REGION Network 16: Actions for STATE Num:49 Wait for Centering Slide Advance
   RUNG wire#powerrail
      Contact( #s49_WaitCentSlideAdv )
      Coil( #qCenteringSlideAdvance )
   END_RUNG
   // the same network as SCL:
   #qCenteringSlideAdvance := #s49_WaitCentSlideAdv;
END_REGION

REGION Network 17: Transition for STATE Num:50 Wait for Distance Sensor Feed Back
   RUNG wire#powerrail
      Contact( #s50_WaitDistSensorFB )
      Contact( #sSst )
      Coil( #s50_WaitDistSensorFB_T1 )
   END_RUNG
   // the same network as SCL:
   #s50_WaitDistSensorFB_T1 := #s50_WaitDistSensorFB AND #sSst;
END_REGION

REGION Network 18: STATE Num:50 Wait for Distance Sensor Feed Back
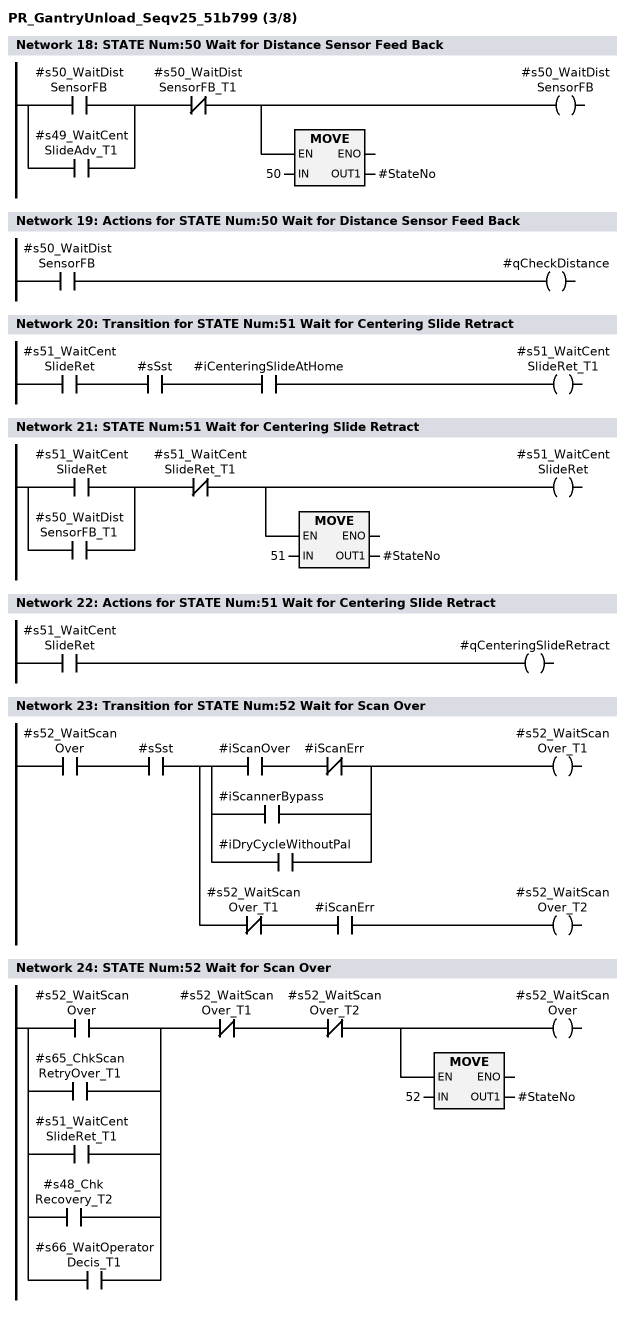
   RUNG wire#powerrail
      Contact( #s50_WaitDistSensorFB )
      wire#w1
      I_Contact( #s50_WaitDistSensorFB_T1 )
      wire#w2
      Coil( #s50_WaitDistSensorFB )
   END_RUNG
   RUNG wire#powerrail
      Contact( #s49_WaitCentSlideAdv_T1 )
   END_RUNG wire#w1
   RUNG wire#w2
      { S7_GenerateENO := "TRUE" } Move(in := 50, out1 => #StateNo)
   END_RUNG
   // the same network as SCL:
   #s50_WaitDistSensorFB := (#s50_WaitDistSensorFB OR #s49_WaitCentSlideAdv_T1) AND NOT #s50_WaitDistSensorFB_T1;
   IF #s50_WaitDistSensorFB THEN #StateNo := 50; END_IF;
END_REGION

REGION Network 19: Actions for STATE Num:50 Wait for Distance Sensor Feed Back
   RUNG wire#powerrail
      Contact( #s50_WaitDistSensorFB )
      Coil( #qCheckDistance )
   END_RUNG
   // the same network as SCL:
   #qCheckDistance := #s50_WaitDistSensorFB;
END_REGION

REGION Network 20: Transition for STATE Num:51 Wait for Centering Slide Retract
   RUNG wire#powerrail
      Contact( #s51_WaitCentSlideRet )
      Contact( #sSst )
      Contact( #iCenteringSlideAtHome )
      Coil( #s51_WaitCentSlideRet_T1 )
   END_RUNG
   // the same network as SCL:
   #s51_WaitCentSlideRet_T1 := #s51_WaitCentSlideRet AND #sSst AND #iCenteringSlideAtHome;
END_REGION

REGION Network 21: STATE Num:51 Wait for Centering Slide Retract
   RUNG wire#powerrail
      Contact( #s51_WaitCentSlideRet )
      wire#w1
      I_Contact( #s51_WaitCentSlideRet_T1 )
      wire#w2
      Coil( #s51_WaitCentSlideRet )
   END_RUNG
   RUNG wire#powerrail
      Contact( #s50_WaitDistSensorFB_T1 )
   END_RUNG wire#w1
   RUNG wire#w2
      { S7_GenerateENO := "TRUE" } Move(in := 51, out1 => #StateNo)
   END_RUNG
   // the same network as SCL:
   #s51_WaitCentSlideRet := (#s51_WaitCentSlideRet OR #s50_WaitDistSensorFB_T1) AND NOT #s51_WaitCentSlideRet_T1;
   IF #s51_WaitCentSlideRet THEN #StateNo := 51; END_IF;
END_REGION

REGION Network 22: Actions for STATE Num:51 Wait for Centering Slide Retract
   RUNG wire#powerrail
      Contact( #s51_WaitCentSlideRet )
      Coil( #qCenteringSlideRetract )
   END_RUNG
   // the same network as SCL:
   #qCenteringSlideRetract := #s51_WaitCentSlideRet;
END_REGION

REGION Network 23: Transition for STATE Num:52 Wait for Scan Over
   RUNG wire#powerrail
      Contact( #s52_WaitScanOver )
      Contact( #sSst )
      wire#w1
      Contact( #iScanOver )
      I_Contact( #iScanErr )
      wire#w2
      Coil( #s52_WaitScanOver_T1 )
   END_RUNG
   RUNG wire#w1
      Contact( #iScannerBypass )
   END_RUNG wire#w2
   RUNG wire#w1
      Contact( #iDryCycleWithoutPal )
   END_RUNG wire#w2
   RUNG wire#w1
      I_Contact( #s52_WaitScanOver_T1 )
      Contact( #iScanErr )
      Coil( #s52_WaitScanOver_T2 )
   END_RUNG
   // the same network as SCL:
   #_w1 := #s52_WaitScanOver AND #sSst;
   #s52_WaitScanOver_T1 := #_w1 AND ((#iScanOver AND NOT #iScanErr) OR #iScannerBypass OR #iDryCycleWithoutPal);
   #s52_WaitScanOver_T2 := #_w1 AND NOT #s52_WaitScanOver_T1 AND #iScanErr;
END_REGION

REGION Network 24: STATE Num:52 Wait for Scan Over
   RUNG wire#powerrail
      Contact( #s52_WaitScanOver )
      wire#w1
      I_Contact( #s52_WaitScanOver_T1 )
      I_Contact( #s52_WaitScanOver_T2 )
      wire#w2
      Coil( #s52_WaitScanOver )
   END_RUNG
   RUNG wire#powerrail
      Contact( #s65_ChkScanRetryOver_T1 )
   END_RUNG wire#w1
   RUNG wire#powerrail
      Contact( #s51_WaitCentSlideRet_T1 )
   END_RUNG wire#w1
   RUNG wire#powerrail
      Contact( #s48_ChkRecovery_T2 )
   END_RUNG wire#w1
   RUNG wire#powerrail
      Contact( #s66_WaitOperatorDecis_T1 )
   END_RUNG wire#w1
   RUNG wire#w2
      { S7_GenerateENO := "TRUE" } Move(in := 52, out1 => #StateNo)
   END_RUNG
   // the same network as SCL:
   #s52_WaitScanOver := (#s52_WaitScanOver OR #s65_ChkScanRetryOver_T1 OR #s51_WaitCentSlideRet_T1 OR #s48_ChkRecovery_T2 OR #s66_WaitOperatorDecis_T1) AND NOT #s52_WaitScanOver_T1 AND NOT #s52_WaitScanOver_T2;
   IF #s52_WaitScanOver THEN #StateNo := 52; END_IF;
END_REGION

REGION Network 25: Actions for STATE Num:52 Wait for Scan Over
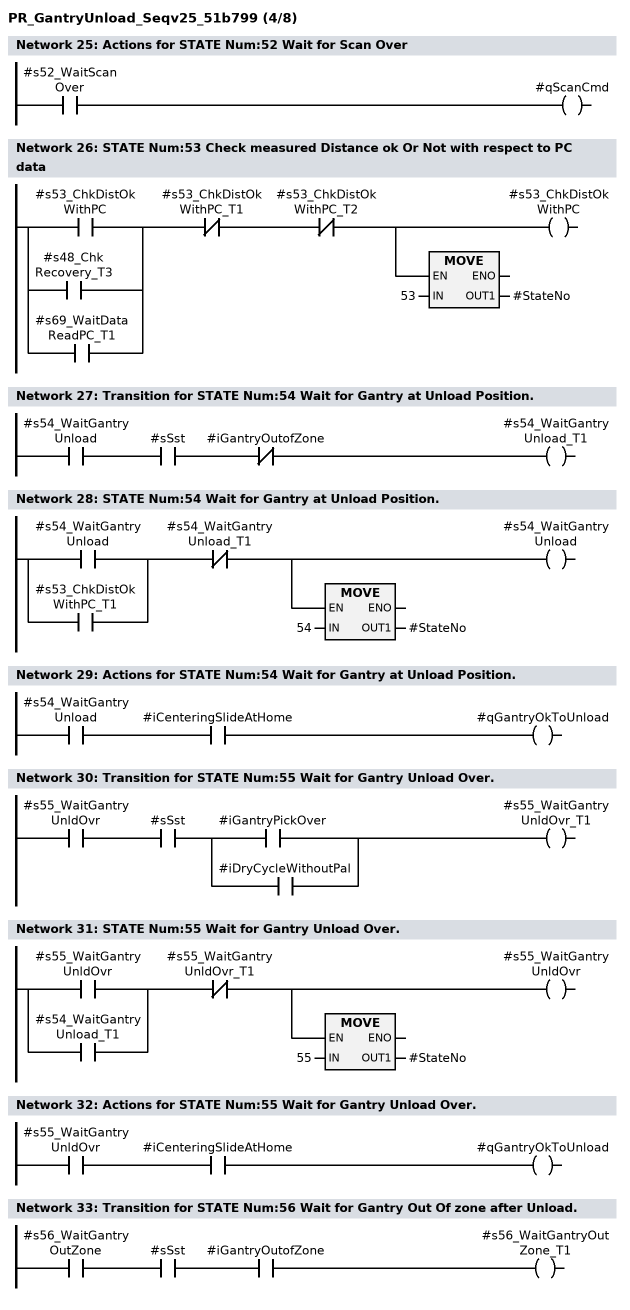
   RUNG wire#powerrail
      Contact( #s52_WaitScanOver )
      Coil( #qScanCmd )
   END_RUNG
   // the same network as SCL:
   #qScanCmd := #s52_WaitScanOver;
END_REGION

REGION Network 26: STATE Num:53 Check measured Distance ok Or Not with respect to PC data
   RUNG wire#powerrail
      Contact( #s53_ChkDistOkWithPC )
      wire#w1
      I_Contact( #s53_ChkDistOkWithPC_T1 )
      I_Contact( #s53_ChkDistOkWithPC_T2 )
      wire#w2
      Coil( #s53_ChkDistOkWithPC )
   END_RUNG
   RUNG wire#powerrail
      Contact( #s48_ChkRecovery_T3 )
   END_RUNG wire#w1
   RUNG wire#powerrail
      Contact( #s69_WaitDataReadPC_T1 )
   END_RUNG wire#w1
   RUNG wire#w2
      { S7_GenerateENO := "TRUE" } Move(in := 53, out1 => #StateNo)
   END_RUNG
   // the same network as SCL:
   #s53_ChkDistOkWithPC := (#s53_ChkDistOkWithPC OR #s48_ChkRecovery_T3 OR #s69_WaitDataReadPC_T1) AND NOT #s53_ChkDistOkWithPC_T1 AND NOT #s53_ChkDistOkWithPC_T2;
   IF #s53_ChkDistOkWithPC THEN #StateNo := 53; END_IF;
END_REGION

REGION Network 27: Transition for STATE Num:54 Wait for Gantry at Unload Position.
   RUNG wire#powerrail
      Contact( #s54_WaitGantryUnload )
      Contact( #sSst )
      I_Contact( #iGantryOutofZone )
      Coil( #s54_WaitGantryUnload_T1 )
   END_RUNG
   // the same network as SCL:
   #s54_WaitGantryUnload_T1 := #s54_WaitGantryUnload AND #sSst AND NOT #iGantryOutofZone;
END_REGION

REGION Network 28: STATE Num:54 Wait for Gantry at Unload Position.
   RUNG wire#powerrail
      Contact( #s54_WaitGantryUnload )
      wire#w1
      I_Contact( #s54_WaitGantryUnload_T1 )
      wire#w2
      Coil( #s54_WaitGantryUnload )
   END_RUNG
   RUNG wire#powerrail
      Contact( #s53_ChkDistOkWithPC_T1 )
   END_RUNG wire#w1
   RUNG wire#w2
      { S7_GenerateENO := "TRUE" } Move(in := 54, out1 => #StateNo)
   END_RUNG
   // the same network as SCL:
   #s54_WaitGantryUnload := (#s54_WaitGantryUnload OR #s53_ChkDistOkWithPC_T1) AND NOT #s54_WaitGantryUnload_T1;
   IF #s54_WaitGantryUnload THEN #StateNo := 54; END_IF;
END_REGION

REGION Network 29: Actions for STATE Num:54 Wait for Gantry at Unload Position.
   RUNG wire#powerrail
      Contact( #s54_WaitGantryUnload )
      Contact( #iCenteringSlideAtHome )
      Coil( #qGantryOkToUnload )
   END_RUNG
   // the same network as SCL:
   #qGantryOkToUnload := #s54_WaitGantryUnload AND #iCenteringSlideAtHome;
END_REGION

REGION Network 30: Transition for STATE Num:55 Wait for Gantry Unload Over.
   RUNG wire#powerrail
      Contact( #s55_WaitGantryUnldOvr )
      Contact( #sSst )
      wire#w1
      Contact( #iGantryPickOver )
      wire#w2
      Coil( #s55_WaitGantryUnldOvr_T1 )
   END_RUNG
   RUNG wire#w1
      Contact( #iDryCycleWithoutPal )
   END_RUNG wire#w2
   // the same network as SCL:
   #s55_WaitGantryUnldOvr_T1 := #s55_WaitGantryUnldOvr AND #sSst AND (#iGantryPickOver OR #iDryCycleWithoutPal);
END_REGION

REGION Network 31: STATE Num:55 Wait for Gantry Unload Over.
   RUNG wire#powerrail
      Contact( #s55_WaitGantryUnldOvr )
      wire#w1
      I_Contact( #s55_WaitGantryUnldOvr_T1 )
      wire#w2
      Coil( #s55_WaitGantryUnldOvr )
   END_RUNG
   RUNG wire#powerrail
      Contact( #s54_WaitGantryUnload_T1 )
   END_RUNG wire#w1
   RUNG wire#w2
      { S7_GenerateENO := "TRUE" } Move(in := 55, out1 => #StateNo)
   END_RUNG
   // the same network as SCL:
   #s55_WaitGantryUnldOvr := (#s55_WaitGantryUnldOvr OR #s54_WaitGantryUnload_T1) AND NOT #s55_WaitGantryUnldOvr_T1;
   IF #s55_WaitGantryUnldOvr THEN #StateNo := 55; END_IF;
END_REGION

REGION Network 32: Actions for STATE Num:55 Wait for Gantry Unload Over.
   RUNG wire#powerrail
      Contact( #s55_WaitGantryUnldOvr )
      Contact( #iCenteringSlideAtHome )
      Coil( #qGantryOkToUnload )
   END_RUNG
   // the same network as SCL:
   #qGantryOkToUnload := #s55_WaitGantryUnldOvr AND #iCenteringSlideAtHome;
END_REGION

REGION Network 33: Transition for STATE Num:56 Wait for Gantry Out Of zone after Unload.
   RUNG wire#powerrail
      Contact( #s56_WaitGantryOutZone )
      Contact( #sSst )
      Contact( #iGantryOutofZone )
      Coil( #s56_WaitGantryOutZone_T1 )
   END_RUNG
   // the same network as SCL:
   #s56_WaitGantryOutZone_T1 := #s56_WaitGantryOutZone AND #sSst AND #iGantryOutofZone;
END_REGION

REGION Network 34: STATE Num:56 Wait for Gantry Out Of zone after Unload.
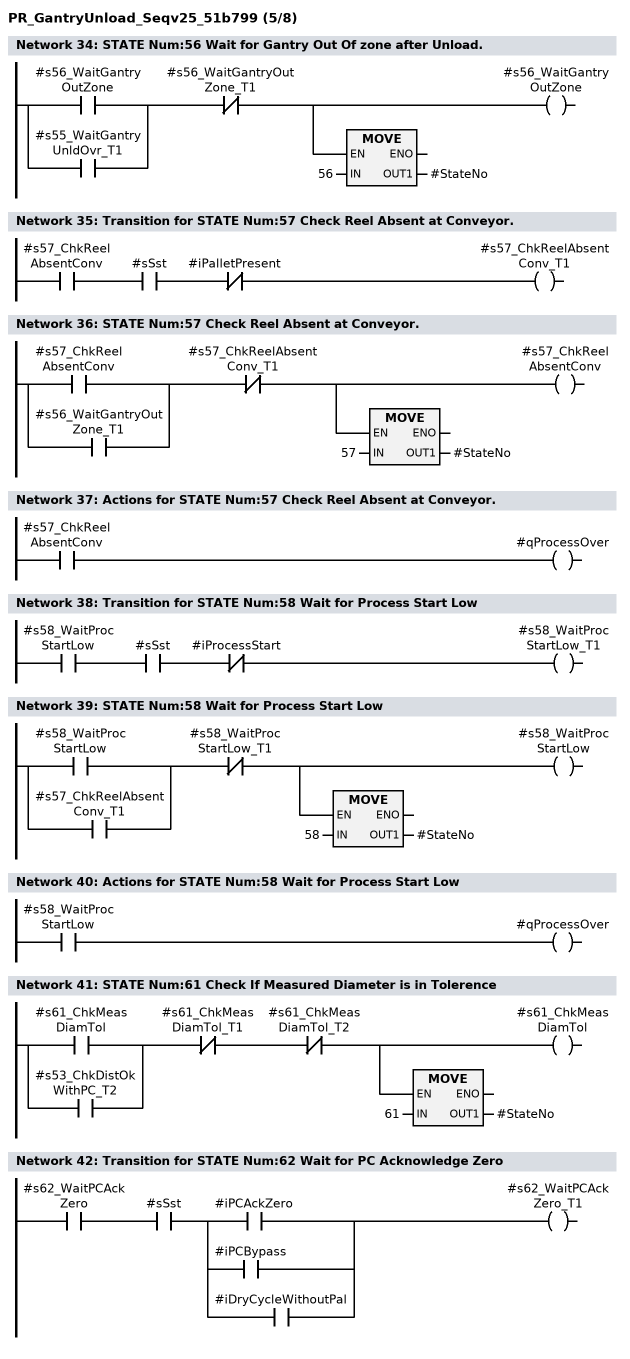
   RUNG wire#powerrail
      Contact( #s56_WaitGantryOutZone )
      wire#w1
      I_Contact( #s56_WaitGantryOutZone_T1 )
      wire#w2
      Coil( #s56_WaitGantryOutZone )
   END_RUNG
   RUNG wire#powerrail
      Contact( #s55_WaitGantryUnldOvr_T1 )
   END_RUNG wire#w1
   RUNG wire#w2
      { S7_GenerateENO := "TRUE" } Move(in := 56, out1 => #StateNo)
   END_RUNG
   // the same network as SCL:
   #s56_WaitGantryOutZone := (#s56_WaitGantryOutZone OR #s55_WaitGantryUnldOvr_T1) AND NOT #s56_WaitGantryOutZone_T1;
   IF #s56_WaitGantryOutZone THEN #StateNo := 56; END_IF;
END_REGION

REGION Network 35: Transition for STATE Num:57 Check Reel Absent at Conveyor.
   RUNG wire#powerrail
      Contact( #s57_ChkReelAbsentConv )
      Contact( #sSst )
      I_Contact( #iPalletPresent )
      Coil( #s57_ChkReelAbsentConv_T1 )
   END_RUNG
   // the same network as SCL:
   #s57_ChkReelAbsentConv_T1 := #s57_ChkReelAbsentConv AND #sSst AND NOT #iPalletPresent;
END_REGION

REGION Network 36: STATE Num:57 Check Reel Absent at Conveyor.
   RUNG wire#powerrail
      Contact( #s57_ChkReelAbsentConv )
      wire#w1
      I_Contact( #s57_ChkReelAbsentConv_T1 )
      wire#w2
      Coil( #s57_ChkReelAbsentConv )
   END_RUNG
   RUNG wire#powerrail
      Contact( #s56_WaitGantryOutZone_T1 )
   END_RUNG wire#w1
   RUNG wire#w2
      { S7_GenerateENO := "TRUE" } Move(in := 57, out1 => #StateNo)
   END_RUNG
   // the same network as SCL:
   #s57_ChkReelAbsentConv := (#s57_ChkReelAbsentConv OR #s56_WaitGantryOutZone_T1) AND NOT #s57_ChkReelAbsentConv_T1;
   IF #s57_ChkReelAbsentConv THEN #StateNo := 57; END_IF;
END_REGION

REGION Network 37: Actions for STATE Num:57 Check Reel Absent at Conveyor.
   RUNG wire#powerrail
      Contact( #s57_ChkReelAbsentConv )
      Coil( #qProcessOver )
   END_RUNG
   // the same network as SCL:
   #qProcessOver := #s57_ChkReelAbsentConv;
END_REGION

REGION Network 38: Transition for STATE Num:58 Wait for Process Start Low
   RUNG wire#powerrail
      Contact( #s58_WaitProcStartLow )
      Contact( #sSst )
      I_Contact( #iProcessStart )
      Coil( #s58_WaitProcStartLow_T1 )
   END_RUNG
   // the same network as SCL:
   #s58_WaitProcStartLow_T1 := #s58_WaitProcStartLow AND #sSst AND NOT #iProcessStart;
END_REGION

REGION Network 39: STATE Num:58 Wait for Process Start Low
   RUNG wire#powerrail
      Contact( #s58_WaitProcStartLow )
      wire#w1
      I_Contact( #s58_WaitProcStartLow_T1 )
      wire#w2
      Coil( #s58_WaitProcStartLow )
   END_RUNG
   RUNG wire#powerrail
      Contact( #s57_ChkReelAbsentConv_T1 )
   END_RUNG wire#w1
   RUNG wire#w2
      { S7_GenerateENO := "TRUE" } Move(in := 58, out1 => #StateNo)
   END_RUNG
   // the same network as SCL:
   #s58_WaitProcStartLow := (#s58_WaitProcStartLow OR #s57_ChkReelAbsentConv_T1) AND NOT #s58_WaitProcStartLow_T1;
   IF #s58_WaitProcStartLow THEN #StateNo := 58; END_IF;
END_REGION

REGION Network 40: Actions for STATE Num:58 Wait for Process Start Low
   RUNG wire#powerrail
      Contact( #s58_WaitProcStartLow )
      Coil( #qProcessOver )
   END_RUNG
   // the same network as SCL:
   #qProcessOver := #s58_WaitProcStartLow;
END_REGION

REGION Network 41: STATE Num:61 Check If Measured Diameter is in Tolerence
   RUNG wire#powerrail
      Contact( #s61_ChkMeasDiamTol )
      wire#w1
      I_Contact( #s61_ChkMeasDiamTol_T1 )
      I_Contact( #s61_ChkMeasDiamTol_T2 )
      wire#w2
      Coil( #s61_ChkMeasDiamTol )
   END_RUNG
   RUNG wire#powerrail
      Contact( #s53_ChkDistOkWithPC_T2 )
   END_RUNG wire#w1
   RUNG wire#w2
      { S7_GenerateENO := "TRUE" } Move(in := 61, out1 => #StateNo)
   END_RUNG
   // the same network as SCL:
   #s61_ChkMeasDiamTol := (#s61_ChkMeasDiamTol OR #s53_ChkDistOkWithPC_T2) AND NOT #s61_ChkMeasDiamTol_T1 AND NOT #s61_ChkMeasDiamTol_T2;
   IF #s61_ChkMeasDiamTol THEN #StateNo := 61; END_IF;
END_REGION

REGION Network 42: Transition for STATE Num:62 Wait for PC Acknowledge Zero
   RUNG wire#powerrail
      Contact( #s62_WaitPCAckZero )
      Contact( #sSst )
      wire#w1
      Contact( #iPCAckZero )
      wire#w2
      Coil( #s62_WaitPCAckZero_T1 )
   END_RUNG
   RUNG wire#w1
      Contact( #iPCBypass )
   END_RUNG wire#w2
   RUNG wire#w1
      Contact( #iDryCycleWithoutPal )
   END_RUNG wire#w2
   // the same network as SCL:
   #s62_WaitPCAckZero_T1 := #s62_WaitPCAckZero AND #sSst AND (#iPCAckZero OR #iPCBypass OR #iDryCycleWithoutPal);
END_REGION

REGION Network 43: STATE Num:62 Wait for PC Acknowledge Zero
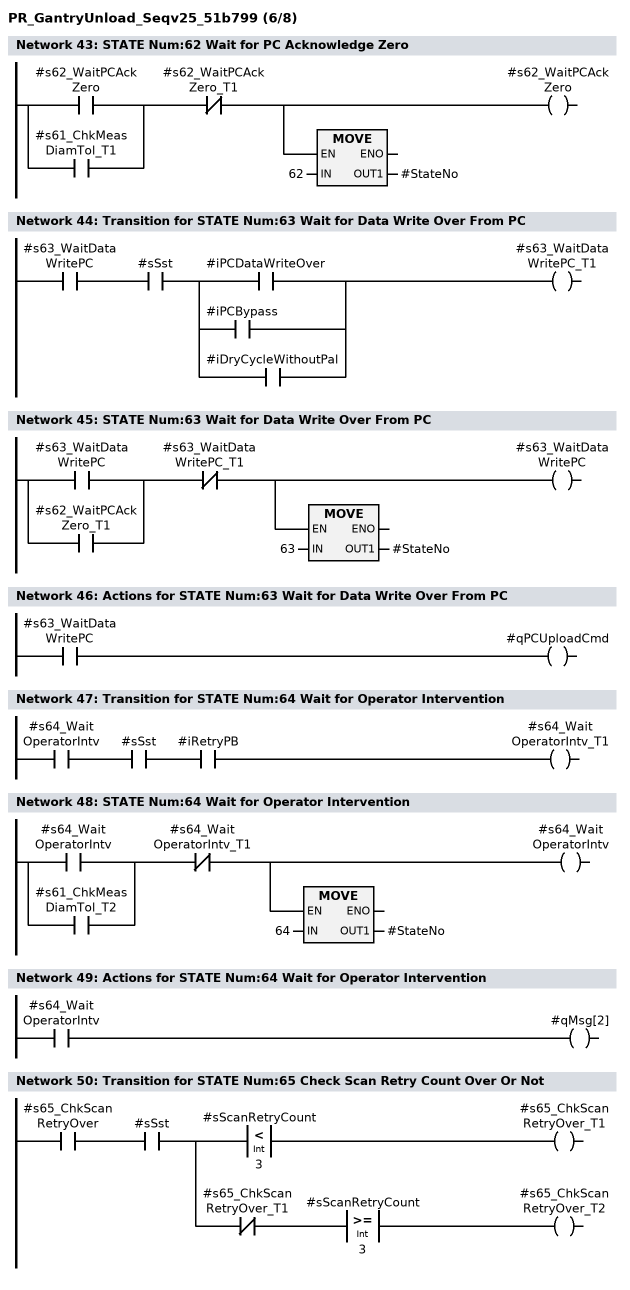
   RUNG wire#powerrail
      Contact( #s62_WaitPCAckZero )
      wire#w1
      I_Contact( #s62_WaitPCAckZero_T1 )
      wire#w2
      Coil( #s62_WaitPCAckZero )
   END_RUNG
   RUNG wire#powerrail
      Contact( #s61_ChkMeasDiamTol_T1 )
   END_RUNG wire#w1
   RUNG wire#w2
      { S7_GenerateENO := "TRUE" } Move(in := 62, out1 => #StateNo)
   END_RUNG
   // the same network as SCL:
   #s62_WaitPCAckZero := (#s62_WaitPCAckZero OR #s61_ChkMeasDiamTol_T1) AND NOT #s62_WaitPCAckZero_T1;
   IF #s62_WaitPCAckZero THEN #StateNo := 62; END_IF;
END_REGION

REGION Network 44: Transition for STATE Num:63 Wait for Data Write Over From PC
   RUNG wire#powerrail
      Contact( #s63_WaitDataWritePC )
      Contact( #sSst )
      wire#w1
      Contact( #iPCDataWriteOver )
      wire#w2
      Coil( #s63_WaitDataWritePC_T1 )
   END_RUNG
   RUNG wire#w1
      Contact( #iPCBypass )
   END_RUNG wire#w2
   RUNG wire#w1
      Contact( #iDryCycleWithoutPal )
   END_RUNG wire#w2
   // the same network as SCL:
   #s63_WaitDataWritePC_T1 := #s63_WaitDataWritePC AND #sSst AND (#iPCDataWriteOver OR #iPCBypass OR #iDryCycleWithoutPal);
END_REGION

REGION Network 45: STATE Num:63 Wait for Data Write Over From PC
   RUNG wire#powerrail
      Contact( #s63_WaitDataWritePC )
      wire#w1
      I_Contact( #s63_WaitDataWritePC_T1 )
      wire#w2
      Coil( #s63_WaitDataWritePC )
   END_RUNG
   RUNG wire#powerrail
      Contact( #s62_WaitPCAckZero_T1 )
   END_RUNG wire#w1
   RUNG wire#w2
      { S7_GenerateENO := "TRUE" } Move(in := 63, out1 => #StateNo)
   END_RUNG
   // the same network as SCL:
   #s63_WaitDataWritePC := (#s63_WaitDataWritePC OR #s62_WaitPCAckZero_T1) AND NOT #s63_WaitDataWritePC_T1;
   IF #s63_WaitDataWritePC THEN #StateNo := 63; END_IF;
END_REGION

REGION Network 46: Actions for STATE Num:63 Wait for Data Write Over From PC
   RUNG wire#powerrail
      Contact( #s63_WaitDataWritePC )
      Coil( #qPCUploadCmd )
   END_RUNG
   // the same network as SCL:
   #qPCUploadCmd := #s63_WaitDataWritePC;
END_REGION

REGION Network 47: Transition for STATE Num:64 Wait for Operator Intervention
   RUNG wire#powerrail
      Contact( #s64_WaitOperatorIntv )
      Contact( #sSst )
      Contact( #iRetryPB )
      Coil( #s64_WaitOperatorIntv_T1 )
   END_RUNG
   // the same network as SCL:
   #s64_WaitOperatorIntv_T1 := #s64_WaitOperatorIntv AND #sSst AND #iRetryPB;
END_REGION

REGION Network 48: STATE Num:64 Wait for Operator Intervention
   RUNG wire#powerrail
      Contact( #s64_WaitOperatorIntv )
      wire#w1
      I_Contact( #s64_WaitOperatorIntv_T1 )
      wire#w2
      Coil( #s64_WaitOperatorIntv )
   END_RUNG
   RUNG wire#powerrail
      Contact( #s61_ChkMeasDiamTol_T2 )
   END_RUNG wire#w1
   RUNG wire#w2
      { S7_GenerateENO := "TRUE" } Move(in := 64, out1 => #StateNo)
   END_RUNG
   // the same network as SCL:
   #s64_WaitOperatorIntv := (#s64_WaitOperatorIntv OR #s61_ChkMeasDiamTol_T2) AND NOT #s64_WaitOperatorIntv_T1;
   IF #s64_WaitOperatorIntv THEN #StateNo := 64; END_IF;
END_REGION

REGION Network 49: Actions for STATE Num:64 Wait for Operator Intervention
   RUNG wire#powerrail
      Contact( #s64_WaitOperatorIntv )
      Coil( #qMsg[2] )
   END_RUNG
   // the same network as SCL:
   #qMsg[2] := #s64_WaitOperatorIntv;
END_REGION

REGION Network 50: Transition for STATE Num:65 Check Scan Retry Count Over Or Not
   RUNG wire#powerrail
      Contact( #s65_ChkScanRetryOver )
      Contact( #sSst )
      wire#w1
      { S7_Templates := "SrcType := Int" } LT_Contact(in1 := #sScanRetryCount, in2 := 3)
      Coil( #s65_ChkScanRetryOver_T1 )
   END_RUNG
   RUNG wire#w1
      I_Contact( #s65_ChkScanRetryOver_T1 )
      { S7_Templates := "SrcType := Int" } GE_Contact(in1 := #sScanRetryCount, in2 := 3)
      Coil( #s65_ChkScanRetryOver_T2 )
   END_RUNG
   // the same network as SCL:
   #_w1 := #s65_ChkScanRetryOver AND #sSst;
   #s65_ChkScanRetryOver_T1 := #_w1 AND (#sScanRetryCount < 3);
   #s65_ChkScanRetryOver_T2 := #_w1 AND NOT #s65_ChkScanRetryOver_T1 AND (#sScanRetryCount >= 3);
END_REGION

REGION Network 51: STATE Num:65 Check Scan Retry Count Over Or Not
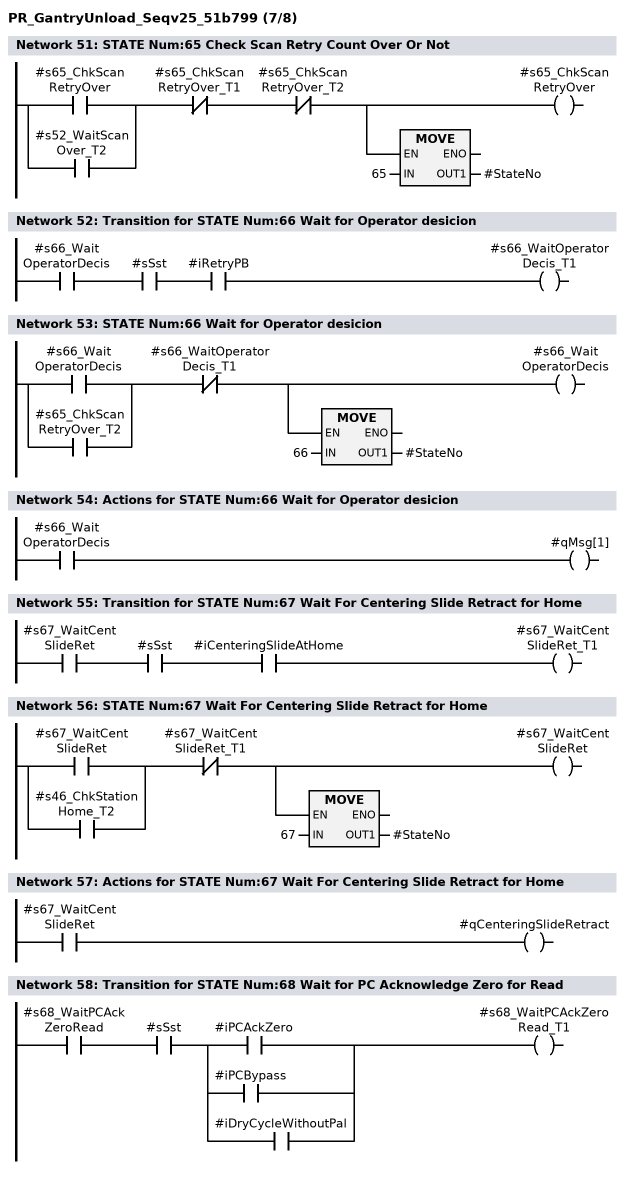
   RUNG wire#powerrail
      Contact( #s65_ChkScanRetryOver )
      wire#w1
      I_Contact( #s65_ChkScanRetryOver_T1 )
      I_Contact( #s65_ChkScanRetryOver_T2 )
      wire#w2
      Coil( #s65_ChkScanRetryOver )
   END_RUNG
   RUNG wire#powerrail
      Contact( #s52_WaitScanOver_T2 )
   END_RUNG wire#w1
   RUNG wire#w2
      { S7_GenerateENO := "TRUE" } Move(in := 65, out1 => #StateNo)
   END_RUNG
   // the same network as SCL:
   #s65_ChkScanRetryOver := (#s65_ChkScanRetryOver OR #s52_WaitScanOver_T2) AND NOT #s65_ChkScanRetryOver_T1 AND NOT #s65_ChkScanRetryOver_T2;
   IF #s65_ChkScanRetryOver THEN #StateNo := 65; END_IF;
END_REGION

REGION Network 52: Transition for STATE Num:66 Wait for Operator desicion
   RUNG wire#powerrail
      Contact( #s66_WaitOperatorDecis )
      Contact( #sSst )
      Contact( #iRetryPB )
      Coil( #s66_WaitOperatorDecis_T1 )
   END_RUNG
   // the same network as SCL:
   #s66_WaitOperatorDecis_T1 := #s66_WaitOperatorDecis AND #sSst AND #iRetryPB;
END_REGION

REGION Network 53: STATE Num:66 Wait for Operator desicion
   RUNG wire#powerrail
      Contact( #s66_WaitOperatorDecis )
      wire#w1
      I_Contact( #s66_WaitOperatorDecis_T1 )
      wire#w2
      Coil( #s66_WaitOperatorDecis )
   END_RUNG
   RUNG wire#powerrail
      Contact( #s65_ChkScanRetryOver_T2 )
   END_RUNG wire#w1
   RUNG wire#w2
      { S7_GenerateENO := "TRUE" } Move(in := 66, out1 => #StateNo)
   END_RUNG
   // the same network as SCL:
   #s66_WaitOperatorDecis := (#s66_WaitOperatorDecis OR #s65_ChkScanRetryOver_T2) AND NOT #s66_WaitOperatorDecis_T1;
   IF #s66_WaitOperatorDecis THEN #StateNo := 66; END_IF;
END_REGION

REGION Network 54: Actions for STATE Num:66 Wait for Operator desicion
   RUNG wire#powerrail
      Contact( #s66_WaitOperatorDecis )
      Coil( #qMsg[1] )
   END_RUNG
   // the same network as SCL:
   #qMsg[1] := #s66_WaitOperatorDecis;
END_REGION

REGION Network 55: Transition for STATE Num:67 Wait For Centering Slide Retract for Home
   RUNG wire#powerrail
      Contact( #s67_WaitCentSlideRet )
      Contact( #sSst )
      Contact( #iCenteringSlideAtHome )
      Coil( #s67_WaitCentSlideRet_T1 )
   END_RUNG
   // the same network as SCL:
   #s67_WaitCentSlideRet_T1 := #s67_WaitCentSlideRet AND #sSst AND #iCenteringSlideAtHome;
END_REGION

REGION Network 56: STATE Num:67 Wait For Centering Slide Retract for Home
   RUNG wire#powerrail
      Contact( #s67_WaitCentSlideRet )
      wire#w1
      I_Contact( #s67_WaitCentSlideRet_T1 )
      wire#w2
      Coil( #s67_WaitCentSlideRet )
   END_RUNG
   RUNG wire#powerrail
      Contact( #s46_ChkStationHome_T2 )
   END_RUNG wire#w1
   RUNG wire#w2
      { S7_GenerateENO := "TRUE" } Move(in := 67, out1 => #StateNo)
   END_RUNG
   // the same network as SCL:
   #s67_WaitCentSlideRet := (#s67_WaitCentSlideRet OR #s46_ChkStationHome_T2) AND NOT #s67_WaitCentSlideRet_T1;
   IF #s67_WaitCentSlideRet THEN #StateNo := 67; END_IF;
END_REGION

REGION Network 57: Actions for STATE Num:67 Wait For Centering Slide Retract for Home
   RUNG wire#powerrail
      Contact( #s67_WaitCentSlideRet )
      Coil( #qCenteringSlideRetract )
   END_RUNG
   // the same network as SCL:
   #qCenteringSlideRetract := #s67_WaitCentSlideRet;
END_REGION

REGION Network 58: Transition for STATE Num:68 Wait for PC Acknowledge Zero for Read
   RUNG wire#powerrail
      Contact( #s68_WaitPCAckZeroRead )
      Contact( #sSst )
      wire#w1
      Contact( #iPCAckZero )
      wire#w2
      Coil( #s68_WaitPCAckZeroRead_T1 )
   END_RUNG
   RUNG wire#w1
      Contact( #iPCBypass )
   END_RUNG wire#w2
   RUNG wire#w1
      Contact( #iDryCycleWithoutPal )
   END_RUNG wire#w2
   // the same network as SCL:
   #s68_WaitPCAckZeroRead_T1 := #s68_WaitPCAckZeroRead AND #sSst AND (#iPCAckZero OR #iPCBypass OR #iDryCycleWithoutPal);
END_REGION

REGION Network 59: STATE Num:68 Wait for PC Acknowledge Zero for Read
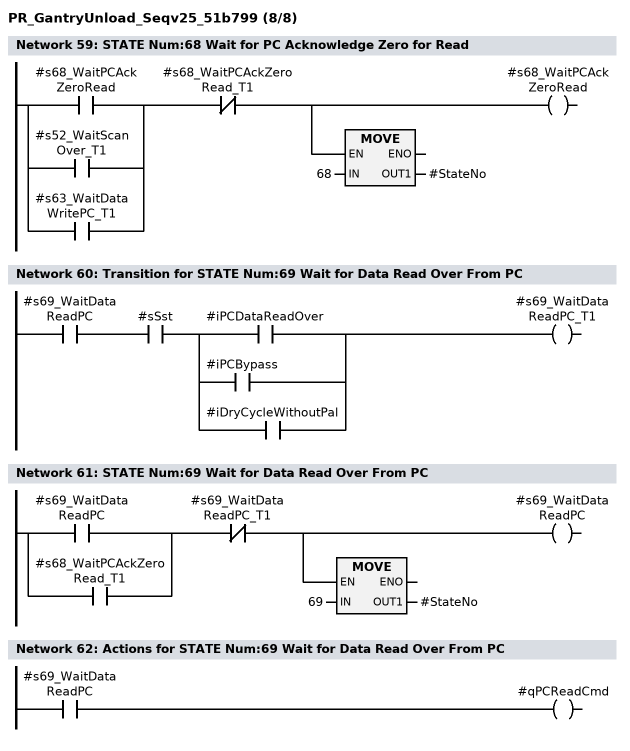
   RUNG wire#powerrail
      Contact( #s68_WaitPCAckZeroRead )
      wire#w1
      I_Contact( #s68_WaitPCAckZeroRead_T1 )
      wire#w2
      Coil( #s68_WaitPCAckZeroRead )
   END_RUNG
   RUNG wire#powerrail
      Contact( #s52_WaitScanOver_T1 )
   END_RUNG wire#w1
   RUNG wire#powerrail
      Contact( #s63_WaitDataWritePC_T1 )
   END_RUNG wire#w1
   RUNG wire#w2
      { S7_GenerateENO := "TRUE" } Move(in := 68, out1 => #StateNo)
   END_RUNG
   // the same network as SCL:
   #s68_WaitPCAckZeroRead := (#s68_WaitPCAckZeroRead OR #s52_WaitScanOver_T1 OR #s63_WaitDataWritePC_T1) AND NOT #s68_WaitPCAckZeroRead_T1;
   IF #s68_WaitPCAckZeroRead THEN #StateNo := 68; END_IF;
END_REGION

REGION Network 60: Transition for STATE Num:69 Wait for Data Read Over From PC
   RUNG wire#powerrail
      Contact( #s69_WaitDataReadPC )
      Contact( #sSst )
      wire#w1
      Contact( #iPCDataReadOver )
      wire#w2
      Coil( #s69_WaitDataReadPC_T1 )
   END_RUNG
   RUNG wire#w1
      Contact( #iPCBypass )
   END_RUNG wire#w2
   RUNG wire#w1
      Contact( #iDryCycleWithoutPal )
   END_RUNG wire#w2
   // the same network as SCL:
   #s69_WaitDataReadPC_T1 := #s69_WaitDataReadPC AND #sSst AND (#iPCDataReadOver OR #iPCBypass OR #iDryCycleWithoutPal);
END_REGION

REGION Network 61: STATE Num:69 Wait for Data Read Over From PC
   RUNG wire#powerrail
      Contact( #s69_WaitDataReadPC )
      wire#w1
      I_Contact( #s69_WaitDataReadPC_T1 )
      wire#w2
      Coil( #s69_WaitDataReadPC )
   END_RUNG
   RUNG wire#powerrail
      Contact( #s68_WaitPCAckZeroRead_T1 )
   END_RUNG wire#w1
   RUNG wire#w2
      { S7_GenerateENO := "TRUE" } Move(in := 69, out1 => #StateNo)
   END_RUNG
   // the same network as SCL:
   #s69_WaitDataReadPC := (#s69_WaitDataReadPC OR #s68_WaitPCAckZeroRead_T1) AND NOT #s69_WaitDataReadPC_T1;
   IF #s69_WaitDataReadPC THEN #StateNo := 69; END_IF;
END_REGION

REGION Network 62: Actions for STATE Num:69 Wait for Data Read Over From PC
   RUNG wire#powerrail
      Contact( #s69_WaitDataReadPC )
      Coil( #qPCReadCmd )
   END_RUNG
   // the same network as SCL:
   #qPCReadCmd := #s69_WaitDataReadPC;
END_REGION
END_FUNCTION_BLOCK

FUNCTION_BLOCK "FB_PR_GantryUnload_Seqv25_V1_V2"   // FB16, LAD
{ S7_Optimized_Access := 'TRUE' }
   VAR_INPUT
      iAutoRunning : Bool;
      iCenteringSlideAtHome : Bool;
      iCenteringSlideAtWork : Bool;
      iDistSenHighLimit : Int;
      iDistSenLowLimit : Int;
      iDistSensorIP : Int;
      iDryCycleWithoutPal : Bool;
      iGantryOutofZone : Bool;
      iGantryPickOver : Bool;
      iPCAckZero : Bool;
      iPCBypass : Bool;
      iPCDataReadOver : Bool;
      iPCDataWriteOver : Bool;
      iPalletPresent : Bool;
      iProcessStart : Bool;
      iReset_fault : Bool;
      iRetryPB : Bool;
      iScanErr : Bool;
      iScanOver : Bool;
      iScannerBypass : Bool;
      iSstMode : Bool;
      iSstPB : Bool;
   END_VAR
   VAR_OUTPUT
      qCenteringSlideAdvance : Bool;
      qCenteringSlideRetract : Bool;
      qCheckDistance : Bool;
      qGantryOkToUnload : Bool;
      qMsg : Array[0..2] of Bool;
      qPCReadCmd : Bool;
      qPCUploadCmd : Bool;
      qProcessOver : Bool;
      qScanCmd : Bool;
   END_VAR
   VAR
      StateNo : Int;
      s44_WaitResetRelease : Bool;
      s44_WaitResetRelease_T1 : Bool;
      s45_WaitGantryOutZone : Bool;
      s45_WaitGantryOutZone_T1 : Bool;
      s46_ChkStationHome : Bool;
      s46_ChkStationHome_T1 : Bool;
      s46_ChkStationHome_T2 : Bool;
      s47_WaitProcStartPZR : Bool;
      s47_WaitProcStartPZR_T1 : Bool;
      s48_ChkRecovery : Bool;
      s48_ChkRecovery_T1 : Bool;
      s48_ChkRecovery_T2 : Bool;
      s48_ChkRecovery_T3 : Bool;
      s49_WaitCentSlideAdv : Bool;
      s49_WaitCentSlideAdv_T1 : Bool;
      s50_WaitDistSensorFB : Bool;
      s50_WaitDistSensorFB_T1 : Bool;
      s51_WaitCentSlideRet : Bool;
      s51_WaitCentSlideRet_T1 : Bool;
      s52_WaitScanOver : Bool;
      s52_WaitScanOver_T1 : Bool;
      s52_WaitScanOver_T2 : Bool;
      s53_ChkMeasDistPCDat : Bool;
      s53_ChkMeasDistPCDat_T1 : Bool;
      s53_ChkMeasDistPCDat_T2 : Bool;
      s54_WaitGantryUnload : Bool;
      s54_WaitGantryUnload_T1 : Bool;
      s55_WaitGantryUnldOvr : Bool;
      s55_WaitGantryUnldOvr_T1 : Bool;
      s56_WaitGantryOutZone : Bool;
      s56_WaitGantryOutZone_T1 : Bool;
      s57_ChkReelAbsentCnv : Bool;
      s57_ChkReelAbsentCnv_T1 : Bool;
      s58_WaitProcStartLow : Bool;
      s58_WaitProcStartLow_T1 : Bool;
      s61_ChkMeasDiamTol : Bool;
      s61_ChkMeasDiamTol_T1 : Bool;
      s61_ChkMeasDiamTol_T2 : Bool;
      s62_WaitPCAckZero : Bool;
      s62_WaitPCAckZero_T1 : Bool;
      s63_WaitDataWritePC : Bool;
      s63_WaitDataWritePC_T1 : Bool;
      s64_WaitOperInterven : Bool;
      s64_WaitOperInterven_T1 : Bool;
      s65_ChkScanRetryOver : Bool;
      s65_ChkScanRetryOver_T1 : Bool;
      s65_ChkScanRetryOver_T2 : Bool;
      s66_WaitOperDecision : Bool;
      s66_WaitOperDecision_T1 : Bool;
      s67_WaitCentSlideRet : Bool;
      s67_WaitCentSlideRet_T1 : Bool;
      s68_WaitPCAckZeroRd : Bool;
      s68_WaitPCAckZeroRd_T1 : Bool;
      s69_WaitDataReadPC : Bool;
      s69_WaitDataReadPC_T1 : Bool;
      sDistanceHighLimit : Int;
      sDistanceLowLimit : Int;
      sRecoveryInt : Int;
      sScanRetryCount : Int;
      sSst : Bool;
      sSstPulse : Bool;
      sSstRise : Bool;
   END_VAR
   VAR_TEMP
      tOne : Bool;
   END_VAR
   VAR_TEMP   // added for the SCL form of the ladder/FBD networks
      _w1 : Bool;
   END_VAR
BEGIN

REGION Network 1
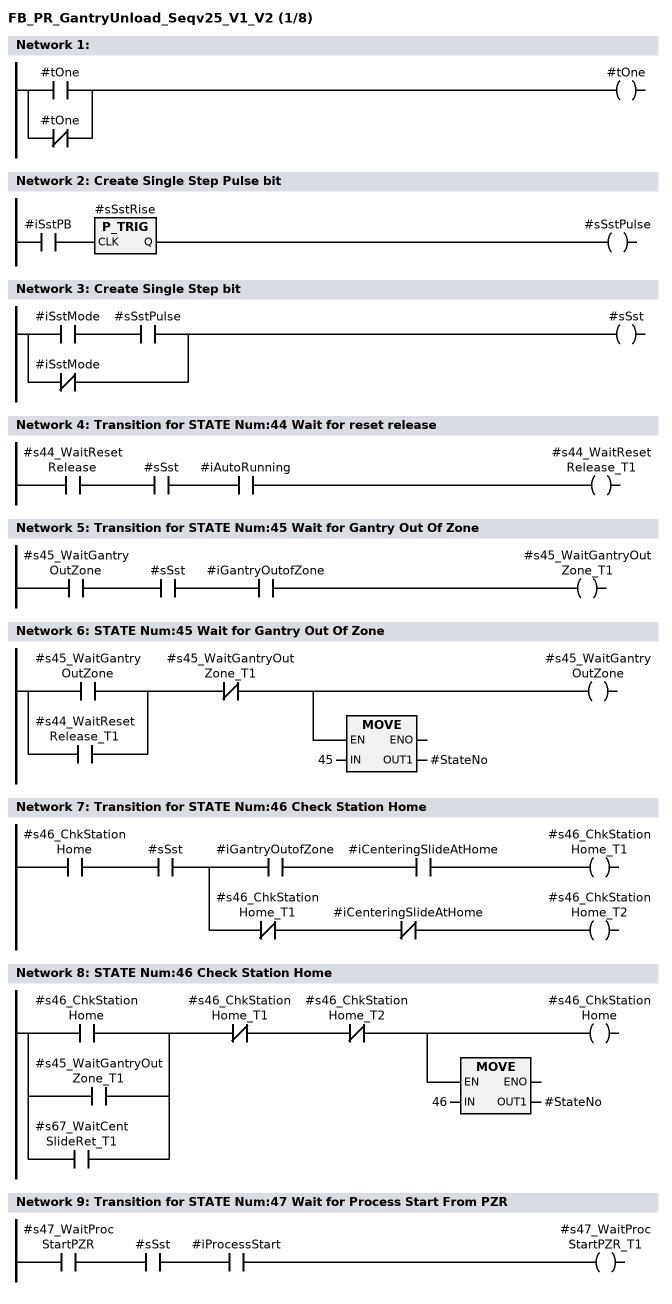
   RUNG wire#powerrail
      Contact( #tOne )
      wire#w1
      Coil( #tOne )
   END_RUNG
   RUNG wire#powerrail
      I_Contact( #tOne )
   END_RUNG wire#w1
   // the same network as SCL:
   #tOne := #tOne OR NOT #tOne;
END_REGION

REGION Network 2: Create Single Step Pulse bit
   RUNG wire#powerrail
      Contact( #iSstPB )
      P_Trig( #sSstRise )
      Coil( #sSstPulse )
   END_RUNG
   // the same network as SCL:
   #_w1 := #iSstPB AND NOT #sSstRise;   // rising edge
   #sSstRise := #iSstPB;
   #sSstPulse := #_w1;
END_REGION

REGION Network 3: Create Single Step bit
   RUNG wire#powerrail
      Contact( #iSstMode )
      Contact( #sSstPulse )
      wire#w1
      Coil( #sSst )
   END_RUNG
   RUNG wire#powerrail
      I_Contact( #iSstMode )
   END_RUNG wire#w1
   // the same network as SCL:
   #sSst := (#iSstMode AND #sSstPulse) OR NOT #iSstMode;
END_REGION

REGION Network 4: Transition for STATE Num:44 Wait for reset release
   RUNG wire#powerrail
      Contact( #s44_WaitResetRelease )
      Contact( #sSst )
      Contact( #iAutoRunning )
      Coil( #s44_WaitResetRelease_T1 )
   END_RUNG
   // the same network as SCL:
   #s44_WaitResetRelease_T1 := #s44_WaitResetRelease AND #sSst AND #iAutoRunning;
END_REGION

REGION Network 5: Transition for STATE Num:45 Wait for Gantry Out Of Zone
   RUNG wire#powerrail
      Contact( #s45_WaitGantryOutZone )
      Contact( #sSst )
      Contact( #iGantryOutofZone )
      Coil( #s45_WaitGantryOutZone_T1 )
   END_RUNG
   // the same network as SCL:
   #s45_WaitGantryOutZone_T1 := #s45_WaitGantryOutZone AND #sSst AND #iGantryOutofZone;
END_REGION

REGION Network 6: STATE Num:45 Wait for Gantry Out Of Zone
   RUNG wire#powerrail
      Contact( #s45_WaitGantryOutZone )
      wire#w1
      I_Contact( #s45_WaitGantryOutZone_T1 )
      wire#w2
      Coil( #s45_WaitGantryOutZone )
   END_RUNG
   RUNG wire#powerrail
      Contact( #s44_WaitResetRelease_T1 )
   END_RUNG wire#w1
   RUNG wire#w2
      { S7_GenerateENO := "TRUE" } Move(in := 45, out1 => #StateNo)
   END_RUNG
   // the same network as SCL:
   #s45_WaitGantryOutZone := (#s45_WaitGantryOutZone OR #s44_WaitResetRelease_T1) AND NOT #s45_WaitGantryOutZone_T1;
   IF #s45_WaitGantryOutZone THEN #StateNo := 45; END_IF;
END_REGION

REGION Network 7: Transition for STATE Num:46 Check Station Home
   RUNG wire#powerrail
      Contact( #s46_ChkStationHome )
      Contact( #sSst )
      wire#w1
      Contact( #iGantryOutofZone )
      Contact( #iCenteringSlideAtHome )
      Coil( #s46_ChkStationHome_T1 )
   END_RUNG
   RUNG wire#w1
      I_Contact( #s46_ChkStationHome_T1 )
      I_Contact( #iCenteringSlideAtHome )
      Coil( #s46_ChkStationHome_T2 )
   END_RUNG
   // the same network as SCL:
   #_w1 := #s46_ChkStationHome AND #sSst;
   #s46_ChkStationHome_T1 := #_w1 AND #iGantryOutofZone AND #iCenteringSlideAtHome;
   #s46_ChkStationHome_T2 := #_w1 AND NOT #s46_ChkStationHome_T1 AND NOT #iCenteringSlideAtHome;
END_REGION

REGION Network 8: STATE Num:46 Check Station Home
   RUNG wire#powerrail
      Contact( #s46_ChkStationHome )
      wire#w1
      I_Contact( #s46_ChkStationHome_T1 )
      I_Contact( #s46_ChkStationHome_T2 )
      wire#w2
      Coil( #s46_ChkStationHome )
   END_RUNG
   RUNG wire#powerrail
      Contact( #s45_WaitGantryOutZone_T1 )
   END_RUNG wire#w1
   RUNG wire#powerrail
      Contact( #s67_WaitCentSlideRet_T1 )
   END_RUNG wire#w1
   RUNG wire#w2
      { S7_GenerateENO := "TRUE" } Move(in := 46, out1 => #StateNo)
   END_RUNG
   // the same network as SCL:
   #s46_ChkStationHome := (#s46_ChkStationHome OR #s45_WaitGantryOutZone_T1 OR #s67_WaitCentSlideRet_T1) AND NOT #s46_ChkStationHome_T1 AND NOT #s46_ChkStationHome_T2;
   IF #s46_ChkStationHome THEN #StateNo := 46; END_IF;
END_REGION

REGION Network 9: Transition for STATE Num:47 Wait for Process Start From PZR
   RUNG wire#powerrail
      Contact( #s47_WaitProcStartPZR )
      Contact( #sSst )
      Contact( #iProcessStart )
      Coil( #s47_WaitProcStartPZR_T1 )
   END_RUNG
   // the same network as SCL:
   #s47_WaitProcStartPZR_T1 := #s47_WaitProcStartPZR AND #sSst AND #iProcessStart;
END_REGION

REGION Network 10: STATE Num:47 Wait for Process Start From PZR
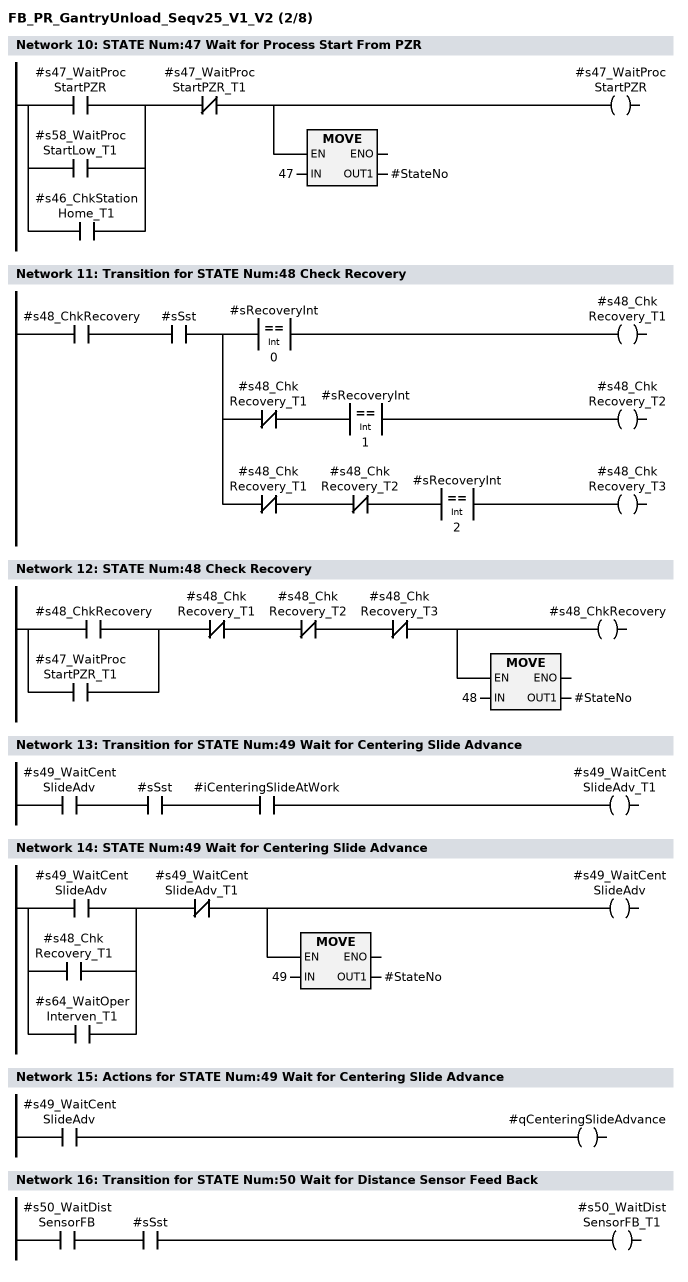
   RUNG wire#powerrail
      Contact( #s47_WaitProcStartPZR )
      wire#w1
      I_Contact( #s47_WaitProcStartPZR_T1 )
      wire#w2
      Coil( #s47_WaitProcStartPZR )
   END_RUNG
   RUNG wire#powerrail
      Contact( #s58_WaitProcStartLow_T1 )
   END_RUNG wire#w1
   RUNG wire#powerrail
      Contact( #s46_ChkStationHome_T1 )
   END_RUNG wire#w1
   RUNG wire#w2
      { S7_GenerateENO := "TRUE" } Move(in := 47, out1 => #StateNo)
   END_RUNG
   // the same network as SCL:
   #s47_WaitProcStartPZR := (#s47_WaitProcStartPZR OR #s58_WaitProcStartLow_T1 OR #s46_ChkStationHome_T1) AND NOT #s47_WaitProcStartPZR_T1;
   IF #s47_WaitProcStartPZR THEN #StateNo := 47; END_IF;
END_REGION

REGION Network 11: Transition for STATE Num:48 Check Recovery
   RUNG wire#powerrail
      Contact( #s48_ChkRecovery )
      Contact( #sSst )
      wire#w1
      { S7_Templates := "SrcType := Int" } EQ_Contact(in1 := #sRecoveryInt, in2 := 0)
      Coil( #s48_ChkRecovery_T1 )
   END_RUNG
   RUNG wire#w1
      I_Contact( #s48_ChkRecovery_T1 )
      { S7_Templates := "SrcType := Int" } EQ_Contact(in1 := #sRecoveryInt, in2 := 1)
      Coil( #s48_ChkRecovery_T2 )
   END_RUNG
   RUNG wire#w1
      I_Contact( #s48_ChkRecovery_T1 )
      I_Contact( #s48_ChkRecovery_T2 )
      { S7_Templates := "SrcType := Int" } EQ_Contact(in1 := #sRecoveryInt, in2 := 2)
      Coil( #s48_ChkRecovery_T3 )
   END_RUNG
   // the same network as SCL:
   #_w1 := #s48_ChkRecovery AND #sSst;
   #s48_ChkRecovery_T1 := #_w1 AND (#sRecoveryInt = 0);
   #s48_ChkRecovery_T2 := #_w1 AND NOT #s48_ChkRecovery_T1 AND (#sRecoveryInt = 1);
   #s48_ChkRecovery_T3 := #_w1 AND NOT #s48_ChkRecovery_T1 AND NOT #s48_ChkRecovery_T2 AND (#sRecoveryInt = 2);
END_REGION

REGION Network 12: STATE Num:48 Check Recovery
   RUNG wire#powerrail
      Contact( #s48_ChkRecovery )
      wire#w1
      I_Contact( #s48_ChkRecovery_T1 )
      I_Contact( #s48_ChkRecovery_T2 )
      I_Contact( #s48_ChkRecovery_T3 )
      wire#w2
      Coil( #s48_ChkRecovery )
   END_RUNG
   RUNG wire#powerrail
      Contact( #s47_WaitProcStartPZR_T1 )
   END_RUNG wire#w1
   RUNG wire#w2
      { S7_GenerateENO := "TRUE" } Move(in := 48, out1 => #StateNo)
   END_RUNG
   // the same network as SCL:
   #s48_ChkRecovery := (#s48_ChkRecovery OR #s47_WaitProcStartPZR_T1) AND NOT #s48_ChkRecovery_T1 AND NOT #s48_ChkRecovery_T2 AND NOT #s48_ChkRecovery_T3;
   IF #s48_ChkRecovery THEN #StateNo := 48; END_IF;
END_REGION

REGION Network 13: Transition for STATE Num:49 Wait for Centering Slide Advance
   RUNG wire#powerrail
      Contact( #s49_WaitCentSlideAdv )
      Contact( #sSst )
      Contact( #iCenteringSlideAtWork )
      Coil( #s49_WaitCentSlideAdv_T1 )
   END_RUNG
   // the same network as SCL:
   #s49_WaitCentSlideAdv_T1 := #s49_WaitCentSlideAdv AND #sSst AND #iCenteringSlideAtWork;
END_REGION

REGION Network 14: STATE Num:49 Wait for Centering Slide Advance
   RUNG wire#powerrail
      Contact( #s49_WaitCentSlideAdv )
      wire#w1
      I_Contact( #s49_WaitCentSlideAdv_T1 )
      wire#w2
      Coil( #s49_WaitCentSlideAdv )
   END_RUNG
   RUNG wire#powerrail
      Contact( #s48_ChkRecovery_T1 )
   END_RUNG wire#w1
   RUNG wire#powerrail
      Contact( #s64_WaitOperInterven_T1 )
   END_RUNG wire#w1
   RUNG wire#w2
      { S7_GenerateENO := "TRUE" } Move(in := 49, out1 => #StateNo)
   END_RUNG
   // the same network as SCL:
   #s49_WaitCentSlideAdv := (#s49_WaitCentSlideAdv OR #s48_ChkRecovery_T1 OR #s64_WaitOperInterven_T1) AND NOT #s49_WaitCentSlideAdv_T1;
   IF #s49_WaitCentSlideAdv THEN #StateNo := 49; END_IF;
END_REGION

REGION Network 15: Actions for STATE Num:49 Wait for Centering Slide Advance
   RUNG wire#powerrail
      Contact( #s49_WaitCentSlideAdv )
      Coil( #qCenteringSlideAdvance )
   END_RUNG
   // the same network as SCL:
   #qCenteringSlideAdvance := #s49_WaitCentSlideAdv;
END_REGION

REGION Network 16: Transition for STATE Num:50 Wait for Distance Sensor Feed Back
   RUNG wire#powerrail
      Contact( #s50_WaitDistSensorFB )
      Contact( #sSst )
      Coil( #s50_WaitDistSensorFB_T1 )
   END_RUNG
   // the same network as SCL:
   #s50_WaitDistSensorFB_T1 := #s50_WaitDistSensorFB AND #sSst;
END_REGION

REGION Network 17: STATE Num:50 Wait for Distance Sensor Feed Back
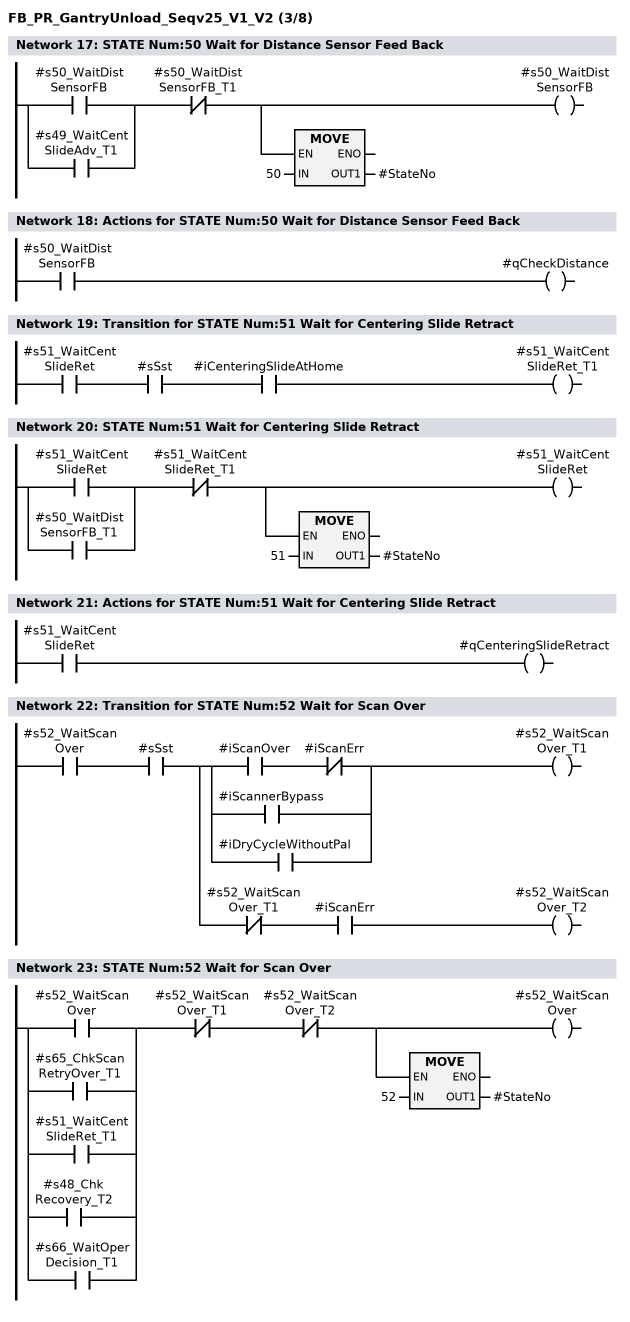
   RUNG wire#powerrail
      Contact( #s50_WaitDistSensorFB )
      wire#w1
      I_Contact( #s50_WaitDistSensorFB_T1 )
      wire#w2
      Coil( #s50_WaitDistSensorFB )
   END_RUNG
   RUNG wire#powerrail
      Contact( #s49_WaitCentSlideAdv_T1 )
   END_RUNG wire#w1
   RUNG wire#w2
      { S7_GenerateENO := "TRUE" } Move(in := 50, out1 => #StateNo)
   END_RUNG
   // the same network as SCL:
   #s50_WaitDistSensorFB := (#s50_WaitDistSensorFB OR #s49_WaitCentSlideAdv_T1) AND NOT #s50_WaitDistSensorFB_T1;
   IF #s50_WaitDistSensorFB THEN #StateNo := 50; END_IF;
END_REGION

REGION Network 18: Actions for STATE Num:50 Wait for Distance Sensor Feed Back
   RUNG wire#powerrail
      Contact( #s50_WaitDistSensorFB )
      Coil( #qCheckDistance )
   END_RUNG
   // the same network as SCL:
   #qCheckDistance := #s50_WaitDistSensorFB;
END_REGION

REGION Network 19: Transition for STATE Num:51 Wait for Centering Slide Retract
   RUNG wire#powerrail
      Contact( #s51_WaitCentSlideRet )
      Contact( #sSst )
      Contact( #iCenteringSlideAtHome )
      Coil( #s51_WaitCentSlideRet_T1 )
   END_RUNG
   // the same network as SCL:
   #s51_WaitCentSlideRet_T1 := #s51_WaitCentSlideRet AND #sSst AND #iCenteringSlideAtHome;
END_REGION

REGION Network 20: STATE Num:51 Wait for Centering Slide Retract
   RUNG wire#powerrail
      Contact( #s51_WaitCentSlideRet )
      wire#w1
      I_Contact( #s51_WaitCentSlideRet_T1 )
      wire#w2
      Coil( #s51_WaitCentSlideRet )
   END_RUNG
   RUNG wire#powerrail
      Contact( #s50_WaitDistSensorFB_T1 )
   END_RUNG wire#w1
   RUNG wire#w2
      { S7_GenerateENO := "TRUE" } Move(in := 51, out1 => #StateNo)
   END_RUNG
   // the same network as SCL:
   #s51_WaitCentSlideRet := (#s51_WaitCentSlideRet OR #s50_WaitDistSensorFB_T1) AND NOT #s51_WaitCentSlideRet_T1;
   IF #s51_WaitCentSlideRet THEN #StateNo := 51; END_IF;
END_REGION

REGION Network 21: Actions for STATE Num:51 Wait for Centering Slide Retract
   RUNG wire#powerrail
      Contact( #s51_WaitCentSlideRet )
      Coil( #qCenteringSlideRetract )
   END_RUNG
   // the same network as SCL:
   #qCenteringSlideRetract := #s51_WaitCentSlideRet;
END_REGION

REGION Network 22: Transition for STATE Num:52 Wait for Scan Over
   RUNG wire#powerrail
      Contact( #s52_WaitScanOver )
      Contact( #sSst )
      wire#w1
      Contact( #iScanOver )
      I_Contact( #iScanErr )
      wire#w2
      Coil( #s52_WaitScanOver_T1 )
   END_RUNG
   RUNG wire#w1
      Contact( #iScannerBypass )
   END_RUNG wire#w2
   RUNG wire#w1
      Contact( #iDryCycleWithoutPal )
   END_RUNG wire#w2
   RUNG wire#w1
      I_Contact( #s52_WaitScanOver_T1 )
      Contact( #iScanErr )
      Coil( #s52_WaitScanOver_T2 )
   END_RUNG
   // the same network as SCL:
   #_w1 := #s52_WaitScanOver AND #sSst;
   #s52_WaitScanOver_T1 := #_w1 AND ((#iScanOver AND NOT #iScanErr) OR #iScannerBypass OR #iDryCycleWithoutPal);
   #s52_WaitScanOver_T2 := #_w1 AND NOT #s52_WaitScanOver_T1 AND #iScanErr;
END_REGION

REGION Network 23: STATE Num:52 Wait for Scan Over
   RUNG wire#powerrail
      Contact( #s52_WaitScanOver )
      wire#w1
      I_Contact( #s52_WaitScanOver_T1 )
      I_Contact( #s52_WaitScanOver_T2 )
      wire#w2
      Coil( #s52_WaitScanOver )
   END_RUNG
   RUNG wire#powerrail
      Contact( #s65_ChkScanRetryOver_T1 )
   END_RUNG wire#w1
   RUNG wire#powerrail
      Contact( #s51_WaitCentSlideRet_T1 )
   END_RUNG wire#w1
   RUNG wire#powerrail
      Contact( #s48_ChkRecovery_T2 )
   END_RUNG wire#w1
   RUNG wire#powerrail
      Contact( #s66_WaitOperDecision_T1 )
   END_RUNG wire#w1
   RUNG wire#w2
      { S7_GenerateENO := "TRUE" } Move(in := 52, out1 => #StateNo)
   END_RUNG
   // the same network as SCL:
   #s52_WaitScanOver := (#s52_WaitScanOver OR #s65_ChkScanRetryOver_T1 OR #s51_WaitCentSlideRet_T1 OR #s48_ChkRecovery_T2 OR #s66_WaitOperDecision_T1) AND NOT #s52_WaitScanOver_T1 AND NOT #s52_WaitScanOver_T2;
   IF #s52_WaitScanOver THEN #StateNo := 52; END_IF;
END_REGION

REGION Network 24: Actions for STATE Num:52 Wait for Scan Over
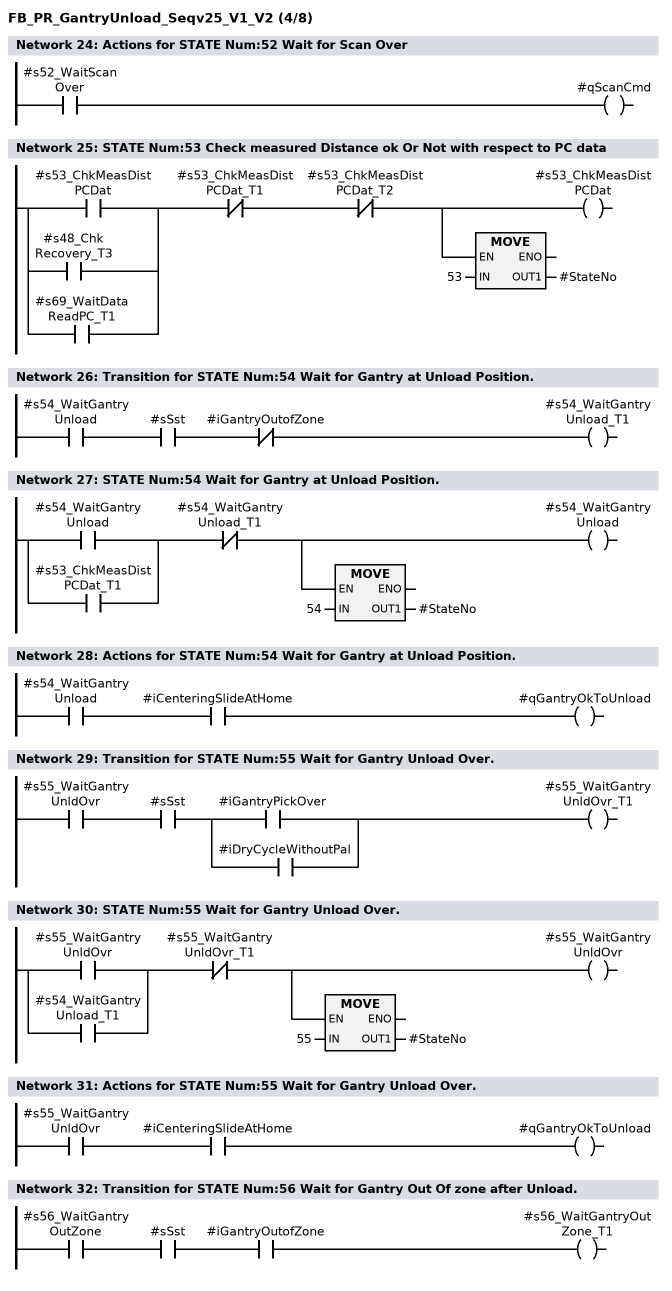
   RUNG wire#powerrail
      Contact( #s52_WaitScanOver )
      Coil( #qScanCmd )
   END_RUNG
   // the same network as SCL:
   #qScanCmd := #s52_WaitScanOver;
END_REGION

REGION Network 25: STATE Num:53 Check measured Distance ok Or Not with respect to PC data
   RUNG wire#powerrail
      Contact( #s53_ChkMeasDistPCDat )
      wire#w1
      I_Contact( #s53_ChkMeasDistPCDat_T1 )
      I_Contact( #s53_ChkMeasDistPCDat_T2 )
      wire#w2
      Coil( #s53_ChkMeasDistPCDat )
   END_RUNG
   RUNG wire#powerrail
      Contact( #s48_ChkRecovery_T3 )
   END_RUNG wire#w1
   RUNG wire#powerrail
      Contact( #s69_WaitDataReadPC_T1 )
   END_RUNG wire#w1
   RUNG wire#w2
      { S7_GenerateENO := "TRUE" } Move(in := 53, out1 => #StateNo)
   END_RUNG
   // the same network as SCL:
   #s53_ChkMeasDistPCDat := (#s53_ChkMeasDistPCDat OR #s48_ChkRecovery_T3 OR #s69_WaitDataReadPC_T1) AND NOT #s53_ChkMeasDistPCDat_T1 AND NOT #s53_ChkMeasDistPCDat_T2;
   IF #s53_ChkMeasDistPCDat THEN #StateNo := 53; END_IF;
END_REGION

REGION Network 26: Transition for STATE Num:54 Wait for Gantry at Unload Position.
   RUNG wire#powerrail
      Contact( #s54_WaitGantryUnload )
      Contact( #sSst )
      I_Contact( #iGantryOutofZone )
      Coil( #s54_WaitGantryUnload_T1 )
   END_RUNG
   // the same network as SCL:
   #s54_WaitGantryUnload_T1 := #s54_WaitGantryUnload AND #sSst AND NOT #iGantryOutofZone;
END_REGION

REGION Network 27: STATE Num:54 Wait for Gantry at Unload Position.
   RUNG wire#powerrail
      Contact( #s54_WaitGantryUnload )
      wire#w1
      I_Contact( #s54_WaitGantryUnload_T1 )
      wire#w2
      Coil( #s54_WaitGantryUnload )
   END_RUNG
   RUNG wire#powerrail
      Contact( #s53_ChkMeasDistPCDat_T1 )
   END_RUNG wire#w1
   RUNG wire#w2
      { S7_GenerateENO := "TRUE" } Move(in := 54, out1 => #StateNo)
   END_RUNG
   // the same network as SCL:
   #s54_WaitGantryUnload := (#s54_WaitGantryUnload OR #s53_ChkMeasDistPCDat_T1) AND NOT #s54_WaitGantryUnload_T1;
   IF #s54_WaitGantryUnload THEN #StateNo := 54; END_IF;
END_REGION

REGION Network 28: Actions for STATE Num:54 Wait for Gantry at Unload Position.
   RUNG wire#powerrail
      Contact( #s54_WaitGantryUnload )
      Contact( #iCenteringSlideAtHome )
      Coil( #qGantryOkToUnload )
   END_RUNG
   // the same network as SCL:
   #qGantryOkToUnload := #s54_WaitGantryUnload AND #iCenteringSlideAtHome;
END_REGION

REGION Network 29: Transition for STATE Num:55 Wait for Gantry Unload Over.
   RUNG wire#powerrail
      Contact( #s55_WaitGantryUnldOvr )
      Contact( #sSst )
      wire#w1
      Contact( #iGantryPickOver )
      wire#w2
      Coil( #s55_WaitGantryUnldOvr_T1 )
   END_RUNG
   RUNG wire#w1
      Contact( #iDryCycleWithoutPal )
   END_RUNG wire#w2
   // the same network as SCL:
   #s55_WaitGantryUnldOvr_T1 := #s55_WaitGantryUnldOvr AND #sSst AND (#iGantryPickOver OR #iDryCycleWithoutPal);
END_REGION

REGION Network 30: STATE Num:55 Wait for Gantry Unload Over.
   RUNG wire#powerrail
      Contact( #s55_WaitGantryUnldOvr )
      wire#w1
      I_Contact( #s55_WaitGantryUnldOvr_T1 )
      wire#w2
      Coil( #s55_WaitGantryUnldOvr )
   END_RUNG
   RUNG wire#powerrail
      Contact( #s54_WaitGantryUnload_T1 )
   END_RUNG wire#w1
   RUNG wire#w2
      { S7_GenerateENO := "TRUE" } Move(in := 55, out1 => #StateNo)
   END_RUNG
   // the same network as SCL:
   #s55_WaitGantryUnldOvr := (#s55_WaitGantryUnldOvr OR #s54_WaitGantryUnload_T1) AND NOT #s55_WaitGantryUnldOvr_T1;
   IF #s55_WaitGantryUnldOvr THEN #StateNo := 55; END_IF;
END_REGION

REGION Network 31: Actions for STATE Num:55 Wait for Gantry Unload Over.
   RUNG wire#powerrail
      Contact( #s55_WaitGantryUnldOvr )
      Contact( #iCenteringSlideAtHome )
      Coil( #qGantryOkToUnload )
   END_RUNG
   // the same network as SCL:
   #qGantryOkToUnload := #s55_WaitGantryUnldOvr AND #iCenteringSlideAtHome;
END_REGION

REGION Network 32: Transition for STATE Num:56 Wait for Gantry Out Of zone after Unload.
   RUNG wire#powerrail
      Contact( #s56_WaitGantryOutZone )
      Contact( #sSst )
      Contact( #iGantryOutofZone )
      Coil( #s56_WaitGantryOutZone_T1 )
   END_RUNG
   // the same network as SCL:
   #s56_WaitGantryOutZone_T1 := #s56_WaitGantryOutZone AND #sSst AND #iGantryOutofZone;
END_REGION

REGION Network 33: STATE Num:56 Wait for Gantry Out Of zone after Unload.
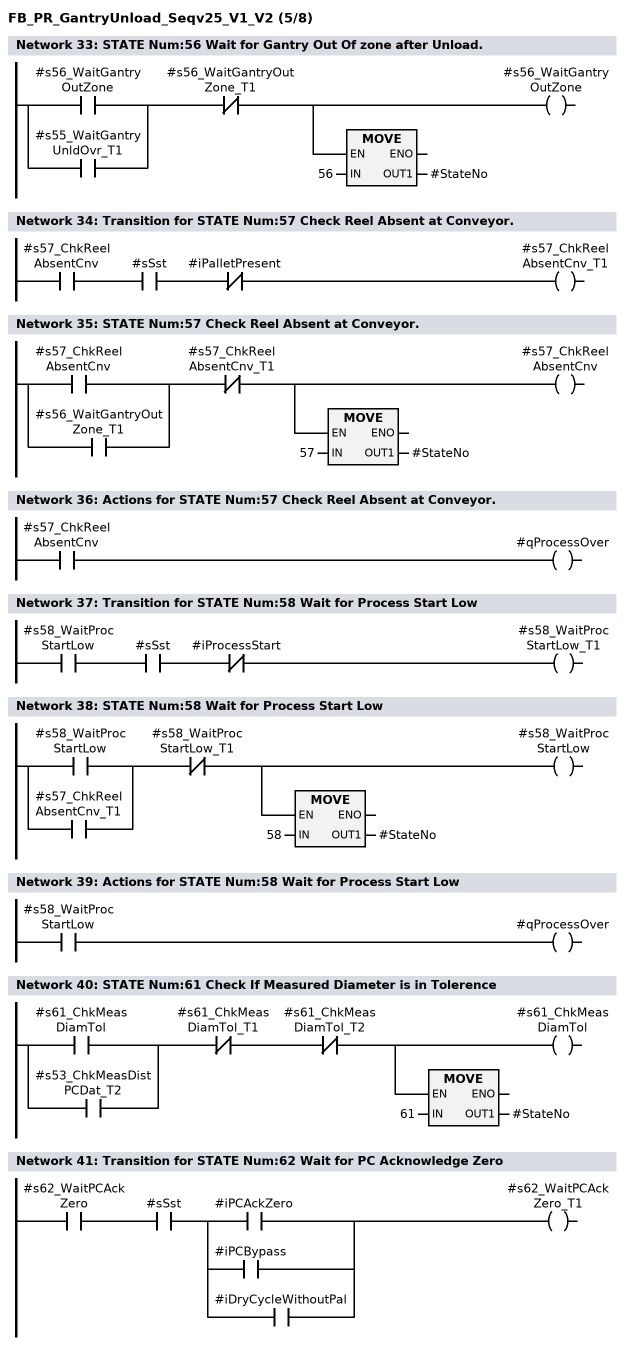
   RUNG wire#powerrail
      Contact( #s56_WaitGantryOutZone )
      wire#w1
      I_Contact( #s56_WaitGantryOutZone_T1 )
      wire#w2
      Coil( #s56_WaitGantryOutZone )
   END_RUNG
   RUNG wire#powerrail
      Contact( #s55_WaitGantryUnldOvr_T1 )
   END_RUNG wire#w1
   RUNG wire#w2
      { S7_GenerateENO := "TRUE" } Move(in := 56, out1 => #StateNo)
   END_RUNG
   // the same network as SCL:
   #s56_WaitGantryOutZone := (#s56_WaitGantryOutZone OR #s55_WaitGantryUnldOvr_T1) AND NOT #s56_WaitGantryOutZone_T1;
   IF #s56_WaitGantryOutZone THEN #StateNo := 56; END_IF;
END_REGION

REGION Network 34: Transition for STATE Num:57 Check Reel Absent at Conveyor.
   RUNG wire#powerrail
      Contact( #s57_ChkReelAbsentCnv )
      Contact( #sSst )
      I_Contact( #iPalletPresent )
      Coil( #s57_ChkReelAbsentCnv_T1 )
   END_RUNG
   // the same network as SCL:
   #s57_ChkReelAbsentCnv_T1 := #s57_ChkReelAbsentCnv AND #sSst AND NOT #iPalletPresent;
END_REGION

REGION Network 35: STATE Num:57 Check Reel Absent at Conveyor.
   RUNG wire#powerrail
      Contact( #s57_ChkReelAbsentCnv )
      wire#w1
      I_Contact( #s57_ChkReelAbsentCnv_T1 )
      wire#w2
      Coil( #s57_ChkReelAbsentCnv )
   END_RUNG
   RUNG wire#powerrail
      Contact( #s56_WaitGantryOutZone_T1 )
   END_RUNG wire#w1
   RUNG wire#w2
      { S7_GenerateENO := "TRUE" } Move(in := 57, out1 => #StateNo)
   END_RUNG
   // the same network as SCL:
   #s57_ChkReelAbsentCnv := (#s57_ChkReelAbsentCnv OR #s56_WaitGantryOutZone_T1) AND NOT #s57_ChkReelAbsentCnv_T1;
   IF #s57_ChkReelAbsentCnv THEN #StateNo := 57; END_IF;
END_REGION

REGION Network 36: Actions for STATE Num:57 Check Reel Absent at Conveyor.
   RUNG wire#powerrail
      Contact( #s57_ChkReelAbsentCnv )
      Coil( #qProcessOver )
   END_RUNG
   // the same network as SCL:
   #qProcessOver := #s57_ChkReelAbsentCnv;
END_REGION

REGION Network 37: Transition for STATE Num:58 Wait for Process Start Low
   RUNG wire#powerrail
      Contact( #s58_WaitProcStartLow )
      Contact( #sSst )
      I_Contact( #iProcessStart )
      Coil( #s58_WaitProcStartLow_T1 )
   END_RUNG
   // the same network as SCL:
   #s58_WaitProcStartLow_T1 := #s58_WaitProcStartLow AND #sSst AND NOT #iProcessStart;
END_REGION

REGION Network 38: STATE Num:58 Wait for Process Start Low
   RUNG wire#powerrail
      Contact( #s58_WaitProcStartLow )
      wire#w1
      I_Contact( #s58_WaitProcStartLow_T1 )
      wire#w2
      Coil( #s58_WaitProcStartLow )
   END_RUNG
   RUNG wire#powerrail
      Contact( #s57_ChkReelAbsentCnv_T1 )
   END_RUNG wire#w1
   RUNG wire#w2
      { S7_GenerateENO := "TRUE" } Move(in := 58, out1 => #StateNo)
   END_RUNG
   // the same network as SCL:
   #s58_WaitProcStartLow := (#s58_WaitProcStartLow OR #s57_ChkReelAbsentCnv_T1) AND NOT #s58_WaitProcStartLow_T1;
   IF #s58_WaitProcStartLow THEN #StateNo := 58; END_IF;
END_REGION

REGION Network 39: Actions for STATE Num:58 Wait for Process Start Low
   RUNG wire#powerrail
      Contact( #s58_WaitProcStartLow )
      Coil( #qProcessOver )
   END_RUNG
   // the same network as SCL:
   #qProcessOver := #s58_WaitProcStartLow;
END_REGION

REGION Network 40: STATE Num:61 Check If Measured Diameter is in Tolerence
   RUNG wire#powerrail
      Contact( #s61_ChkMeasDiamTol )
      wire#w1
      I_Contact( #s61_ChkMeasDiamTol_T1 )
      I_Contact( #s61_ChkMeasDiamTol_T2 )
      wire#w2
      Coil( #s61_ChkMeasDiamTol )
   END_RUNG
   RUNG wire#powerrail
      Contact( #s53_ChkMeasDistPCDat_T2 )
   END_RUNG wire#w1
   RUNG wire#w2
      { S7_GenerateENO := "TRUE" } Move(in := 61, out1 => #StateNo)
   END_RUNG
   // the same network as SCL:
   #s61_ChkMeasDiamTol := (#s61_ChkMeasDiamTol OR #s53_ChkMeasDistPCDat_T2) AND NOT #s61_ChkMeasDiamTol_T1 AND NOT #s61_ChkMeasDiamTol_T2;
   IF #s61_ChkMeasDiamTol THEN #StateNo := 61; END_IF;
END_REGION

REGION Network 41: Transition for STATE Num:62 Wait for PC Acknowledge Zero
   RUNG wire#powerrail
      Contact( #s62_WaitPCAckZero )
      Contact( #sSst )
      wire#w1
      Contact( #iPCAckZero )
      wire#w2
      Coil( #s62_WaitPCAckZero_T1 )
   END_RUNG
   RUNG wire#w1
      Contact( #iPCBypass )
   END_RUNG wire#w2
   RUNG wire#w1
      Contact( #iDryCycleWithoutPal )
   END_RUNG wire#w2
   // the same network as SCL:
   #s62_WaitPCAckZero_T1 := #s62_WaitPCAckZero AND #sSst AND (#iPCAckZero OR #iPCBypass OR #iDryCycleWithoutPal);
END_REGION

REGION Network 42: STATE Num:62 Wait for PC Acknowledge Zero
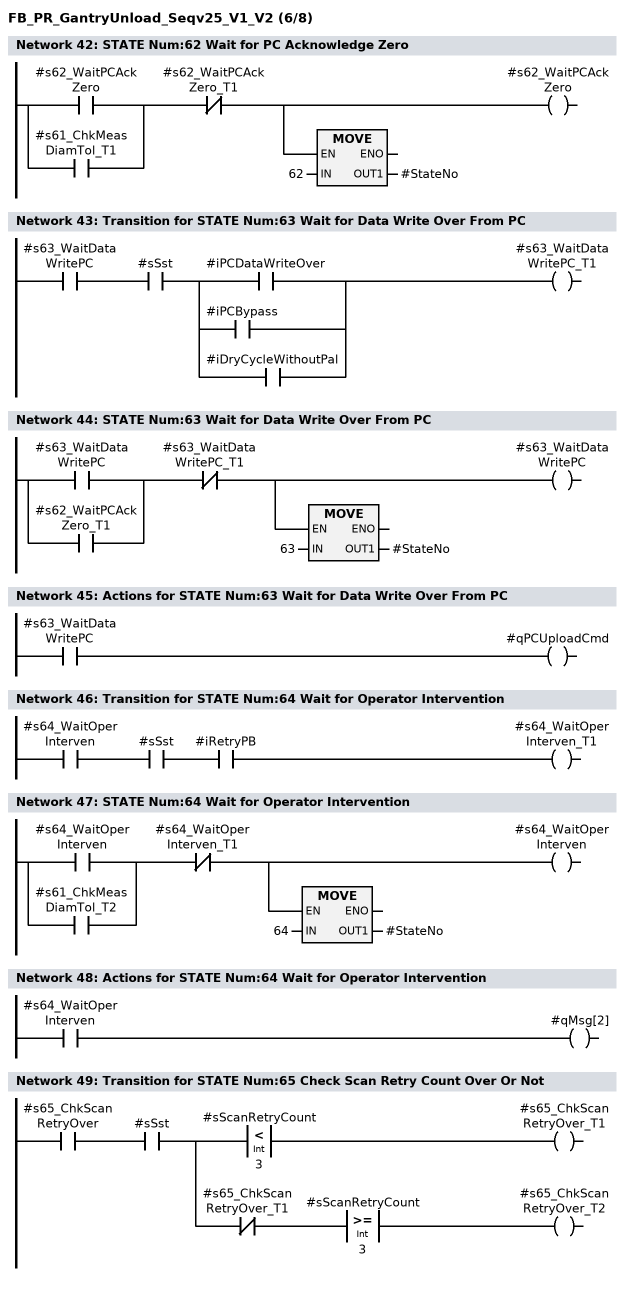
   RUNG wire#powerrail
      Contact( #s62_WaitPCAckZero )
      wire#w1
      I_Contact( #s62_WaitPCAckZero_T1 )
      wire#w2
      Coil( #s62_WaitPCAckZero )
   END_RUNG
   RUNG wire#powerrail
      Contact( #s61_ChkMeasDiamTol_T1 )
   END_RUNG wire#w1
   RUNG wire#w2
      { S7_GenerateENO := "TRUE" } Move(in := 62, out1 => #StateNo)
   END_RUNG
   // the same network as SCL:
   #s62_WaitPCAckZero := (#s62_WaitPCAckZero OR #s61_ChkMeasDiamTol_T1) AND NOT #s62_WaitPCAckZero_T1;
   IF #s62_WaitPCAckZero THEN #StateNo := 62; END_IF;
END_REGION

REGION Network 43: Transition for STATE Num:63 Wait for Data Write Over From PC
   RUNG wire#powerrail
      Contact( #s63_WaitDataWritePC )
      Contact( #sSst )
      wire#w1
      Contact( #iPCDataWriteOver )
      wire#w2
      Coil( #s63_WaitDataWritePC_T1 )
   END_RUNG
   RUNG wire#w1
      Contact( #iPCBypass )
   END_RUNG wire#w2
   RUNG wire#w1
      Contact( #iDryCycleWithoutPal )
   END_RUNG wire#w2
   // the same network as SCL:
   #s63_WaitDataWritePC_T1 := #s63_WaitDataWritePC AND #sSst AND (#iPCDataWriteOver OR #iPCBypass OR #iDryCycleWithoutPal);
END_REGION

REGION Network 44: STATE Num:63 Wait for Data Write Over From PC
   RUNG wire#powerrail
      Contact( #s63_WaitDataWritePC )
      wire#w1
      I_Contact( #s63_WaitDataWritePC_T1 )
      wire#w2
      Coil( #s63_WaitDataWritePC )
   END_RUNG
   RUNG wire#powerrail
      Contact( #s62_WaitPCAckZero_T1 )
   END_RUNG wire#w1
   RUNG wire#w2
      { S7_GenerateENO := "TRUE" } Move(in := 63, out1 => #StateNo)
   END_RUNG
   // the same network as SCL:
   #s63_WaitDataWritePC := (#s63_WaitDataWritePC OR #s62_WaitPCAckZero_T1) AND NOT #s63_WaitDataWritePC_T1;
   IF #s63_WaitDataWritePC THEN #StateNo := 63; END_IF;
END_REGION

REGION Network 45: Actions for STATE Num:63 Wait for Data Write Over From PC
   RUNG wire#powerrail
      Contact( #s63_WaitDataWritePC )
      Coil( #qPCUploadCmd )
   END_RUNG
   // the same network as SCL:
   #qPCUploadCmd := #s63_WaitDataWritePC;
END_REGION

REGION Network 46: Transition for STATE Num:64 Wait for Operator Intervention
   RUNG wire#powerrail
      Contact( #s64_WaitOperInterven )
      Contact( #sSst )
      Contact( #iRetryPB )
      Coil( #s64_WaitOperInterven_T1 )
   END_RUNG
   // the same network as SCL:
   #s64_WaitOperInterven_T1 := #s64_WaitOperInterven AND #sSst AND #iRetryPB;
END_REGION

REGION Network 47: STATE Num:64 Wait for Operator Intervention
   RUNG wire#powerrail
      Contact( #s64_WaitOperInterven )
      wire#w1
      I_Contact( #s64_WaitOperInterven_T1 )
      wire#w2
      Coil( #s64_WaitOperInterven )
   END_RUNG
   RUNG wire#powerrail
      Contact( #s61_ChkMeasDiamTol_T2 )
   END_RUNG wire#w1
   RUNG wire#w2
      { S7_GenerateENO := "TRUE" } Move(in := 64, out1 => #StateNo)
   END_RUNG
   // the same network as SCL:
   #s64_WaitOperInterven := (#s64_WaitOperInterven OR #s61_ChkMeasDiamTol_T2) AND NOT #s64_WaitOperInterven_T1;
   IF #s64_WaitOperInterven THEN #StateNo := 64; END_IF;
END_REGION

REGION Network 48: Actions for STATE Num:64 Wait for Operator Intervention
   RUNG wire#powerrail
      Contact( #s64_WaitOperInterven )
      Coil( #qMsg[2] )
   END_RUNG
   // the same network as SCL:
   #qMsg[2] := #s64_WaitOperInterven;
END_REGION

REGION Network 49: Transition for STATE Num:65 Check Scan Retry Count Over Or Not
   RUNG wire#powerrail
      Contact( #s65_ChkScanRetryOver )
      Contact( #sSst )
      wire#w1
      { S7_Templates := "SrcType := Int" } LT_Contact(in1 := #sScanRetryCount, in2 := 3)
      Coil( #s65_ChkScanRetryOver_T1 )
   END_RUNG
   RUNG wire#w1
      I_Contact( #s65_ChkScanRetryOver_T1 )
      { S7_Templates := "SrcType := Int" } GE_Contact(in1 := #sScanRetryCount, in2 := 3)
      Coil( #s65_ChkScanRetryOver_T2 )
   END_RUNG
   // the same network as SCL:
   #_w1 := #s65_ChkScanRetryOver AND #sSst;
   #s65_ChkScanRetryOver_T1 := #_w1 AND (#sScanRetryCount < 3);
   #s65_ChkScanRetryOver_T2 := #_w1 AND NOT #s65_ChkScanRetryOver_T1 AND (#sScanRetryCount >= 3);
END_REGION

REGION Network 50: STATE Num:65 Check Scan Retry Count Over Or Not
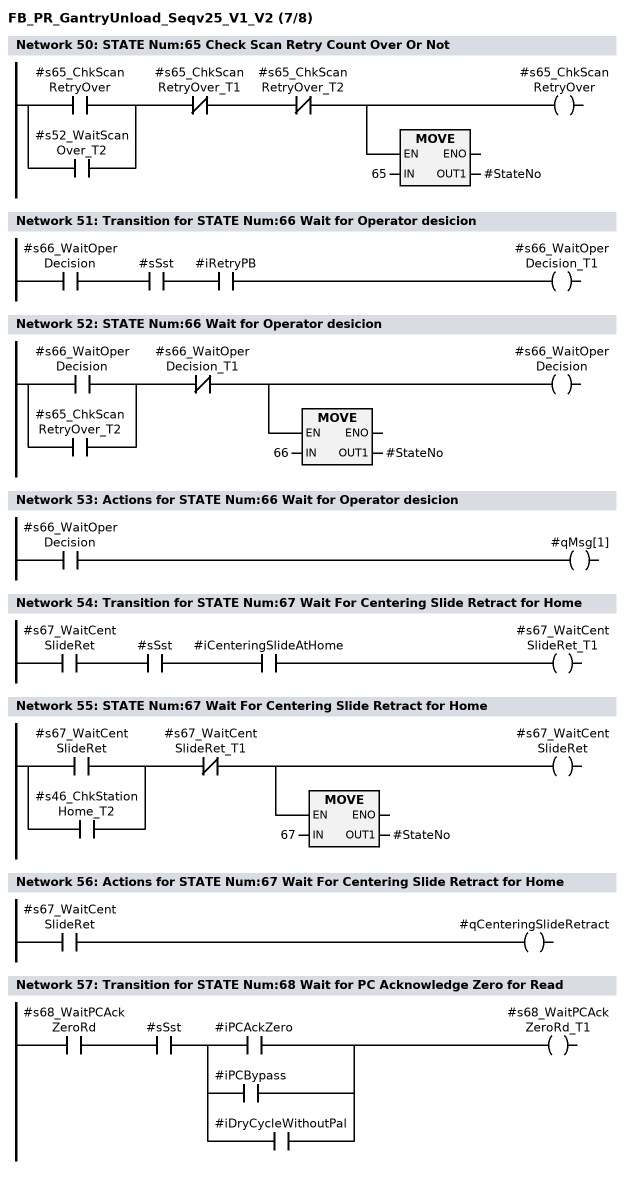
   RUNG wire#powerrail
      Contact( #s65_ChkScanRetryOver )
      wire#w1
      I_Contact( #s65_ChkScanRetryOver_T1 )
      I_Contact( #s65_ChkScanRetryOver_T2 )
      wire#w2
      Coil( #s65_ChkScanRetryOver )
   END_RUNG
   RUNG wire#powerrail
      Contact( #s52_WaitScanOver_T2 )
   END_RUNG wire#w1
   RUNG wire#w2
      { S7_GenerateENO := "TRUE" } Move(in := 65, out1 => #StateNo)
   END_RUNG
   // the same network as SCL:
   #s65_ChkScanRetryOver := (#s65_ChkScanRetryOver OR #s52_WaitScanOver_T2) AND NOT #s65_ChkScanRetryOver_T1 AND NOT #s65_ChkScanRetryOver_T2;
   IF #s65_ChkScanRetryOver THEN #StateNo := 65; END_IF;
END_REGION

REGION Network 51: Transition for STATE Num:66 Wait for Operator desicion
   RUNG wire#powerrail
      Contact( #s66_WaitOperDecision )
      Contact( #sSst )
      Contact( #iRetryPB )
      Coil( #s66_WaitOperDecision_T1 )
   END_RUNG
   // the same network as SCL:
   #s66_WaitOperDecision_T1 := #s66_WaitOperDecision AND #sSst AND #iRetryPB;
END_REGION

REGION Network 52: STATE Num:66 Wait for Operator desicion
   RUNG wire#powerrail
      Contact( #s66_WaitOperDecision )
      wire#w1
      I_Contact( #s66_WaitOperDecision_T1 )
      wire#w2
      Coil( #s66_WaitOperDecision )
   END_RUNG
   RUNG wire#powerrail
      Contact( #s65_ChkScanRetryOver_T2 )
   END_RUNG wire#w1
   RUNG wire#w2
      { S7_GenerateENO := "TRUE" } Move(in := 66, out1 => #StateNo)
   END_RUNG
   // the same network as SCL:
   #s66_WaitOperDecision := (#s66_WaitOperDecision OR #s65_ChkScanRetryOver_T2) AND NOT #s66_WaitOperDecision_T1;
   IF #s66_WaitOperDecision THEN #StateNo := 66; END_IF;
END_REGION

REGION Network 53: Actions for STATE Num:66 Wait for Operator desicion
   RUNG wire#powerrail
      Contact( #s66_WaitOperDecision )
      Coil( #qMsg[1] )
   END_RUNG
   // the same network as SCL:
   #qMsg[1] := #s66_WaitOperDecision;
END_REGION

REGION Network 54: Transition for STATE Num:67 Wait For Centering Slide Retract for Home
   RUNG wire#powerrail
      Contact( #s67_WaitCentSlideRet )
      Contact( #sSst )
      Contact( #iCenteringSlideAtHome )
      Coil( #s67_WaitCentSlideRet_T1 )
   END_RUNG
   // the same network as SCL:
   #s67_WaitCentSlideRet_T1 := #s67_WaitCentSlideRet AND #sSst AND #iCenteringSlideAtHome;
END_REGION

REGION Network 55: STATE Num:67 Wait For Centering Slide Retract for Home
   RUNG wire#powerrail
      Contact( #s67_WaitCentSlideRet )
      wire#w1
      I_Contact( #s67_WaitCentSlideRet_T1 )
      wire#w2
      Coil( #s67_WaitCentSlideRet )
   END_RUNG
   RUNG wire#powerrail
      Contact( #s46_ChkStationHome_T2 )
   END_RUNG wire#w1
   RUNG wire#w2
      { S7_GenerateENO := "TRUE" } Move(in := 67, out1 => #StateNo)
   END_RUNG
   // the same network as SCL:
   #s67_WaitCentSlideRet := (#s67_WaitCentSlideRet OR #s46_ChkStationHome_T2) AND NOT #s67_WaitCentSlideRet_T1;
   IF #s67_WaitCentSlideRet THEN #StateNo := 67; END_IF;
END_REGION

REGION Network 56: Actions for STATE Num:67 Wait For Centering Slide Retract for Home
   RUNG wire#powerrail
      Contact( #s67_WaitCentSlideRet )
      Coil( #qCenteringSlideRetract )
   END_RUNG
   // the same network as SCL:
   #qCenteringSlideRetract := #s67_WaitCentSlideRet;
END_REGION

REGION Network 57: Transition for STATE Num:68 Wait for PC Acknowledge Zero for Read
   RUNG wire#powerrail
      Contact( #s68_WaitPCAckZeroRd )
      Contact( #sSst )
      wire#w1
      Contact( #iPCAckZero )
      wire#w2
      Coil( #s68_WaitPCAckZeroRd_T1 )
   END_RUNG
   RUNG wire#w1
      Contact( #iPCBypass )
   END_RUNG wire#w2
   RUNG wire#w1
      Contact( #iDryCycleWithoutPal )
   END_RUNG wire#w2
   // the same network as SCL:
   #s68_WaitPCAckZeroRd_T1 := #s68_WaitPCAckZeroRd AND #sSst AND (#iPCAckZero OR #iPCBypass OR #iDryCycleWithoutPal);
END_REGION

REGION Network 58: STATE Num:68 Wait for PC Acknowledge Zero for Read
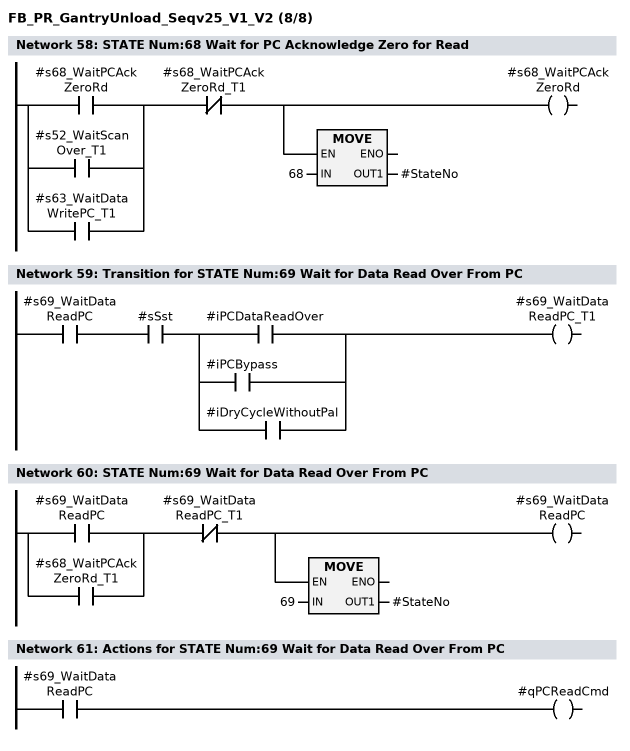
   RUNG wire#powerrail
      Contact( #s68_WaitPCAckZeroRd )
      wire#w1
      I_Contact( #s68_WaitPCAckZeroRd_T1 )
      wire#w2
      Coil( #s68_WaitPCAckZeroRd )
   END_RUNG
   RUNG wire#powerrail
      Contact( #s52_WaitScanOver_T1 )
   END_RUNG wire#w1
   RUNG wire#powerrail
      Contact( #s63_WaitDataWritePC_T1 )
   END_RUNG wire#w1
   RUNG wire#w2
      { S7_GenerateENO := "TRUE" } Move(in := 68, out1 => #StateNo)
   END_RUNG
   // the same network as SCL:
   #s68_WaitPCAckZeroRd := (#s68_WaitPCAckZeroRd OR #s52_WaitScanOver_T1 OR #s63_WaitDataWritePC_T1) AND NOT #s68_WaitPCAckZeroRd_T1;
   IF #s68_WaitPCAckZeroRd THEN #StateNo := 68; END_IF;
END_REGION

REGION Network 59: Transition for STATE Num:69 Wait for Data Read Over From PC
   RUNG wire#powerrail
      Contact( #s69_WaitDataReadPC )
      Contact( #sSst )
      wire#w1
      Contact( #iPCDataReadOver )
      wire#w2
      Coil( #s69_WaitDataReadPC_T1 )
   END_RUNG
   RUNG wire#w1
      Contact( #iPCBypass )
   END_RUNG wire#w2
   RUNG wire#w1
      Contact( #iDryCycleWithoutPal )
   END_RUNG wire#w2
   // the same network as SCL:
   #s69_WaitDataReadPC_T1 := #s69_WaitDataReadPC AND #sSst AND (#iPCDataReadOver OR #iPCBypass OR #iDryCycleWithoutPal);
END_REGION

REGION Network 60: STATE Num:69 Wait for Data Read Over From PC
   RUNG wire#powerrail
      Contact( #s69_WaitDataReadPC )
      wire#w1
      I_Contact( #s69_WaitDataReadPC_T1 )
      wire#w2
      Coil( #s69_WaitDataReadPC )
   END_RUNG
   RUNG wire#powerrail
      Contact( #s68_WaitPCAckZeroRd_T1 )
   END_RUNG wire#w1
   RUNG wire#w2
      { S7_GenerateENO := "TRUE" } Move(in := 69, out1 => #StateNo)
   END_RUNG
   // the same network as SCL:
   #s69_WaitDataReadPC := (#s69_WaitDataReadPC OR #s68_WaitPCAckZeroRd_T1) AND NOT #s69_WaitDataReadPC_T1;
   IF #s69_WaitDataReadPC THEN #StateNo := 69; END_IF;
END_REGION

REGION Network 61: Actions for STATE Num:69 Wait for Data Read Over From PC
   RUNG wire#powerrail
      Contact( #s69_WaitDataReadPC )
      Coil( #qPCReadCmd )
   END_RUNG
   // the same network as SCL:
   #qPCReadCmd := #s69_WaitDataReadPC;
END_REGION
END_FUNCTION_BLOCK

ORGANIZATION_BLOCK "Main"   // OB1, LAD, ProgramCycle
TITLE = "Main Program Sweep (Cycle)"
{ S7_Optimized_Access := 'TRUE' }
VERSION : 0.1
   VAR_INPUT
      Initial_Call : Bool;   // Initial call of this OB
      Remanence : Bool;   // =True, if remanent data are available
   END_VAR
   VAR_TEMP
      OB1_EV_CLASS : Byte;   // Bits 0-3 = 1 (Coming event), Bits 4-7 = 1 (Event class 1)
      OB1_SCAN_1 : Byte;   // 1 (Cold restart scan 1 of OB 1), 3 (Scan 2-n of OB 1)
      OB1_PRIORITY : Byte;   // Priority of OB Execution
      OB1_OB_NUMBR : Byte;   // 1 (Organization block 1, OB1)
      OB1_RESERVED_1 : Byte;   // Reserved for system
      OB1_RESERVED_2 : Byte;   // Reserved for system
      OB1_PREV_CYCLE : Int;   // Cycle time of previous OB1 scan (milliseconds)
      OB1_MIN_CYCLE : Int;   // Minimum cycle time of OB1 (milliseconds)
      OB1_MAX_CYCLE : Int;   // Maximum cycle time of OB1 (milliseconds)
      OB1_DATE_TIME : Date_And_Time;   // Date and time OB1 started
   END_VAR
BEGIN
END_ORGANIZATION_BLOCK

// ===== library types =====

// folder: S2-Process Function Unit

FUNCTION_BLOCK "PR_CognexISCamera_Profinet"   // FB365, LAD
TITLE = Cognex2D_4Feature / Cognex Camera Module
{ S7_Optimized_Access := 'TRUE' }
AUTHOR : Deepak.Jagtap
FAMILY : WIPROPARI
NAME : S21006022005
VERSION : 0.1
// |============================================================================|
// BLOCK:Cognex Camera Module
// Item Code : SMxxxxx
// Owner:Precision Automation & Robotics India Ltd.
// Author: DJ
// Release Date:04-04-2018
// Version:0.1
// V0.1-Initial release
// |============================================================================|
// Block Description: This block is used for interface of Cognex Camera via 
// profinet  and enter Job selection from outside the block.
// |============================================================================|
// Errors:
// qErrTriggerTimeOut: Trigger TimeOut Error Occured
// qErrAcquiringTimeout: Acquiring TimeOut Error Occured
// qErrTriggerEnableTimeout: Trigger Enable TimeOut Occured
// qErrJobSelection: Job selection Error
// qBothStartOn: Both Start are ON
// ============================================================================|
// Dependency:
// Map Vision Input and Output from External IO address. Byte should be matched as per the block
// |============================================================================|
   VAR_INPUT
      iResetFault : Bool;   // Reset Fault Input
      iAutorunning : Bool;   // Autorunning Input
      iStartJobSelection : Bool;   // start job selection / Start for Job Selection
      iStartInspection : Bool;   // Start for Inspection / start inspection
      iRetryCount : Int;   // Retry Count eg:3,4 etc / retry count
      iRetryPB : Bool;
      iJobID : Int;   // Enter Job ID / job id
      iTriggerEnableTimeoutTime : Time;   // Trigger Enable TimeOut Time Delay
      iTriggerTimeoutTime : Time;   // Trigger TimeOut Time Delay
      iAcquiringTimeOutTime : Time;   // Acquiring TimeOut Time Delay
   END_VAR
   VAR_OUTPUT
      qJobPass : Bool;   // Job Pass In Inspection
      qJobFail : Bool;   // Job Failed In Inspection
      qJobSelectionOver : Bool;   // Connect Job Selection over bit / job selection over
      qJobInspectionOver : Bool;   // Inspection Over Output
      qVisionOnline : Bool;   // Insight Vision Is In Online
      qVisionOfflineReason1 : Bool;   // Insight Vision Offline Due To: The vision system's job is being modified
      qVisionOfflineReason2 : Bool;   // Insight Vision Offline Due To: A discrete signal is holding the vision system Offline
      qVisionOfflineReason3 : Bool;   // Insight Vision Offline Due To: A communications protocol is holding the vision system Offline
      qErrBothStartOn : Bool;   // Both Start are On / both start on
      qErrJobSelection : Bool;   // Job selection Error Occur / error job selection
      qErrTriggerEnableTimeout : Bool;   // Trigger Enable TimeOut Error
      qErrTriggerTimeOut : Bool;   // Trigger TimeOut Error
      qErrAcquiringTimeOut : Bool;   // Acquiring TimeOut Error
   END_VAR
   VAR_IN_OUT
      iqInputAddrs : ANY;   // Input HW Address P#I120.0 BYTE 74
      iqOutputAddrs : ANY;   // Input HW Address P#Q120.0 BYTE 68
      iqRetryCount : Int;   // Retry Count Display / Retry count
      iqRunningJobID : Int;   // Running job ID
      iqInsight_Camera : Struct   // Insight Camera PZD
         Vision_Input : Struct
            "iTrigger Ready" : Bool;
            "iTrigger Ack" : Bool;
            iExposureComplete : Bool;
            "iMissed Ack" : Bool;
            "iOffline Reason_0" : Bool;
            "iOffline Reason_1" : Bool;
            "iOffline Reason_2" : Bool;
            iOnline : Bool;
            Acquisition_ID : Byte;
            Acquisition_ID_1 : Byte;
            iSystemBusy : Bool;
            "iInspection Completed" : Bool;
            "iResults Buffer Overrun" : Bool;
            "iResults Valid" : Bool;
            iCommandExecuting : Bool;
            iCommandComplete : Bool;
            "iCommand Failed" : Bool;
            iSetUserDataAck : Bool;
            iJobPass : Bool;
            iReserved : Bool;
            iReserved_1 : Bool;
            iReserved_2 : Bool;
            iReserved_3 : Bool;
            iReserved_4 : Bool;
            iReserved_5 : Bool;
            iError : Bool;
            iErrorCode : Int;
            iCommandControlInput : Int;
            SoftEventControlInput : Byte;
            iInspection_ID : Byte;
            iInspection_ID_1 : Byte;
            iInspection_ResultCode : Byte;
            iInspection_ResultCode_1 : Byte;
            iInspection_Result : Array[213..277] of Byte;
         END_STRUCT;
         Vision_Output : Struct
            "qTrigger Enable" : Bool;
            qTrigger : Bool;
            qClearExposureComplete : Bool;
            qReserved_1 : Bool;
            qReserved_2 : Bool;
            qReserved_3 : Bool;
            qReserved_4 : Bool;
            "qSet Offline" : Bool;
            "qBuffer Results Enable" : Bool;
            "qInspection Results Ack" : Bool;
            qSetUserData : Bool;
            qExecuteCommand : Bool;
            qReserved : Bool;
            qReserved_5 : Bool;
            qReserved_6 : Bool;
            qClearError : Bool;
            qCommandControl : Word;
            "Soft Event Control" : Byte;
            qUser_Data : Array[205..268] of Byte;
         END_STRUCT;
      END_STRUCT;
   END_VAR
   VAR
      sResetFaults : Bool;   // Reset Faults
      sInspectionComplete : Bool;   // Inspection Complete
      TriggerTimeout : TON_TIME;   // TriggerTimeout Timer
      TriggerEnableTimeout : TON_TIME;   // TriggerEnableTimeout Timer
      AcquiringTimeOut : TON_TIME;   // AcquiringTimeOut Timer
      ResultTimer : TON_TIME;   // ResultTimer
      sPulse : Array[0..11] of Bool;   // Array of Pulses
      sJobPass : Bool;   // Stat Bit of Job Pass
      sVisionInputCmdControlIP : Int;
      sJobFail : Bool;   // Stat Bit of Job Fail
      sJobLoadcompleted : Bool;
      sErrTriggerTimeOut : Bool;   // Error Trigger Time Out
      sErrJobSelection : Bool;
      sBothStartOn : Bool;
      sJobSelectionOver : Bool;
      sJobInspectionOver : Bool;
      sErrAcquiringTimeOut : Bool;   // Error Acquiring Time Out
      sErrTriggerEnableTimeout : Bool;   // Error Trigger Enable Time Out
      sVisionOutput_Trigger : Bool;   // Vision Outpur Trigger
      sRetryCountOver : Bool;
      sInitialPulse : Bool;
      sProgramEcho : TON_TIME;
      sExposureTimerStar1 : Bool;
      sExposureTimerStart : Bool;
      sExposureTimer : TON_TIME;
      sExecDelayTimer : TON_TIME;
      sRetry : TON_TIME;
   END_VAR
   VAR_TEMP
      tInspectionID : Int;
      tResultCode : Int;
   END_VAR
   VAR_TEMP   // added for the SCL form of the ladder/FBD networks
      _w1 : Bool;
      _w2 : Bool;
      _w3 : Bool;
      _w4 : Bool;
   END_VAR
BEGIN

REGION Network 1: Header
   // ==============================================================================
   //  Company: Precision Automation & Robotics India Ltd. 
   // ------------------------------------------------------------------------------
   //  Item Code: S21006022005
   //  Author/Created by: Deepak.Jagtap
   //  Reviewed/Checked by: Atul P
   //  First Release on: 04-04-2018
   //  Latest update on:
   // ------------------------------------------------------------------------------
   //  Tested with: CPU firmware, model or simulator testing
   //  Engineering/Editor: TIA Portal V15.1
   // ------------------------------------------------------------------------------
   //  Restrictions:
   //  Dependencies/Requirements:
   // iqInsight_Camera	Struct
   // Map Vision Input and Output from with External IO address
   // ------------------------------------------------------------------------------
   //  Change Log:
   //  Ver.	Date		Changed by		Details of changes
   //  1.0	04-04-2018	Deepak.Jagtap            	First release version
   // 
   // ------------------------------------------------------------------------------
   //  Functionality: This block is used for interface of Cognex Camera via 
   // profinet.
   // 
   //  Inputs
   // iResetFault	Bool
   // iAutorunning	Bool
   // iStartJobSelection	Bool
   // iStartInspection	Bool
   // iRetryCount	Int
   // iJobID	Int
   // iTriggerEnableTimeoutTime	Time
   // iTriggerTimeoutTime	Time
   // iAcquiringTimeOutTime	Time
   // 
   //  Outputs
   // qJobPass	Bool
   // qJobFail	Bool
   // qJobSelectionOver	Bool
   // qJobInspectionOver	Bool
   // qVisionOnline	Bool
   // qVisionOfflineReason1	Bool
   // qVisionOfflineReason2	Bool
   // qVisionOfflineReason3	Bool
   // qErrBothStartOn	Bool
   // qErrJobSelection	Bool
   // qErrTriggerEnableTimeout	Bool
   // qErrTriggerTimeOut	Bool
   // qErrAcquiringTimeOut	Bool
   // 
   //  In-outs
   // iqInputAddrs	Any
   // iqOutputAddrs	Any
   // iqRetryCount	Int
   // iqRunningJobID	Int
   // iqInsight_Camera	Struct
   // 
   // ------------------------------------------------------------------------------
   //  Errors reported:
   //  1.qErrTriggerTimeOut : Error trigger timeout
   // 2. qErrAcquiringTimeOut;Acquiring Time Out
   // 3. qErrTriggerEnableTimeout:Trigger Enable Time Out
   // 4. qErrBothStartOn:both start on
   // 5. qErrJobSelection:error job selection
   //  Messages reported:
   //  1. Message 1 present
   //  2. Message 2 present
   // ==============================================================================
END_REGION

REGION Network 2: Read Data From Input Area
   // Read Data From Input Area
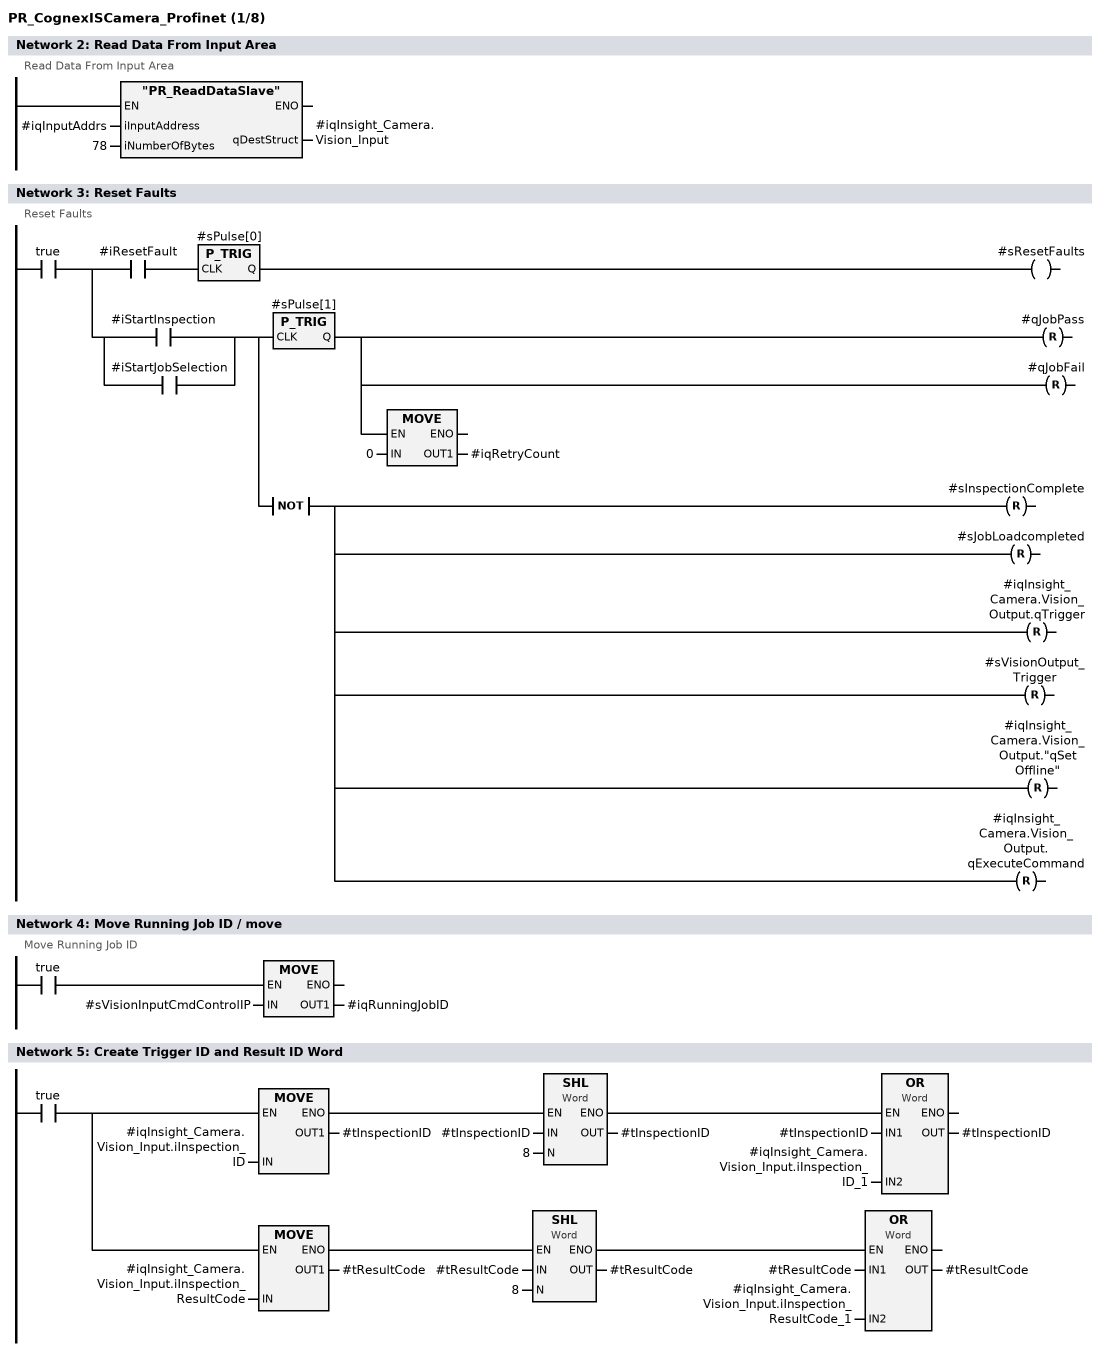
   RUNG wire#powerrail
      "PR_ReadDataSlave"(iInputAddress := #iqInputAddrs, iNumberOfBytes := 78, qDestStruct => #iqInsight_Camera.Vision_Input)
   END_RUNG
   // the same network as SCL:
   "PR_ReadDataSlave"(iInputAddress := #iqInputAddrs,
                      iNumberOfBytes := 78,
                      qDestStruct => #iqInsight_Camera.Vision_Input);
END_REGION

REGION Network 3: Reset Faults
   // Reset Faults
   RUNG wire#powerrail
      Contact( true )
      wire#w1
      Contact( #iResetFault )
      P_Trig( #sPulse[0] )
      Coil( #sResetFaults )
   END_RUNG
   RUNG wire#w1
      Contact( #iStartInspection )
      wire#w2
      P_Trig( #sPulse[1] )
      wire#w3
      R_Coil( #qJobPass )
   END_RUNG
   RUNG wire#w1
      Contact( #iStartJobSelection )
   END_RUNG wire#w2
   RUNG wire#w3
      R_Coil( #qJobFail )
   END_RUNG
   RUNG wire#w3
      Move(in := 0, out1 => #iqRetryCount)
   END_RUNG
   RUNG wire#w2
      Not()
      wire#w4
      R_Coil( #sInspectionComplete )
   END_RUNG
   RUNG wire#w4
      R_Coil( #sJobLoadcompleted )
   END_RUNG
   RUNG wire#w4
      R_Coil( #iqInsight_Camera.Vision_Output.qTrigger )
   END_RUNG
   RUNG wire#w4
      R_Coil( #sVisionOutput_Trigger )
   END_RUNG
   RUNG wire#w4
      R_Coil( #iqInsight_Camera.Vision_Output."qSet Offline" )
   END_RUNG
   RUNG wire#w4
      R_Coil( #iqInsight_Camera.Vision_Output.qExecuteCommand )
   END_RUNG
   // the same network as SCL:
   #_w1 := true AND #iResetFault;
   #_w2 := #_w1 AND NOT #sPulse[0];   // rising edge
   #sPulse[0] := #_w1;
   #sResetFaults := #_w2;
   #_w3 := true AND (#iStartInspection OR #iStartJobSelection);
   #_w4 := #_w3 AND NOT #sPulse[1];   // rising edge
   #sPulse[1] := #_w3;
   IF #_w4 THEN
       #qJobPass := FALSE;
       #qJobFail := FALSE;
       #iqRetryCount := 0;
   END_IF;
   IF NOT #_w3 THEN
       #sInspectionComplete := FALSE;
       #sJobLoadcompleted := FALSE;
       #iqInsight_Camera.Vision_Output.qTrigger := FALSE;
       #sVisionOutput_Trigger := FALSE;
       #iqInsight_Camera.Vision_Output."qSet Offline" := FALSE;
       #iqInsight_Camera.Vision_Output.qExecuteCommand := FALSE;
   END_IF;
END_REGION

REGION Network 4: Move Running Job ID / move
   // Move Running Job ID
   RUNG wire#powerrail
      Contact( true )
      Move(in := #sVisionInputCmdControlIP, out1 => #iqRunningJobID)
   END_RUNG
   // the same network as SCL:
   IF true THEN #iqRunningJobID := #sVisionInputCmdControlIP; END_IF;
END_REGION

REGION Network 5: Create Trigger ID and Result ID Word
   IF true THEN
       #tInspectionID := #iqInsight_Camera.Vision_Input.iInspection_ID;
       #tInspectionID := SHL(IN := #tInspectionID, N := 8);
       #tInspectionID := #tInspectionID OR #iqInsight_Camera.Vision_Input.iInspection_ID_1;
       #tResultCode := #iqInsight_Camera.Vision_Input.iInspection_ResultCode;
       #tResultCode := SHL(IN := #tResultCode, N := 8);
       #tResultCode := #tResultCode OR #iqInsight_Camera.Vision_Input.iInspection_ResultCode_1;
   END_IF;
END_REGION

REGION Network 6: Trigger Enable through Job Selection / Camera Trigger Enable
   // Trigger Enable through Job Selection
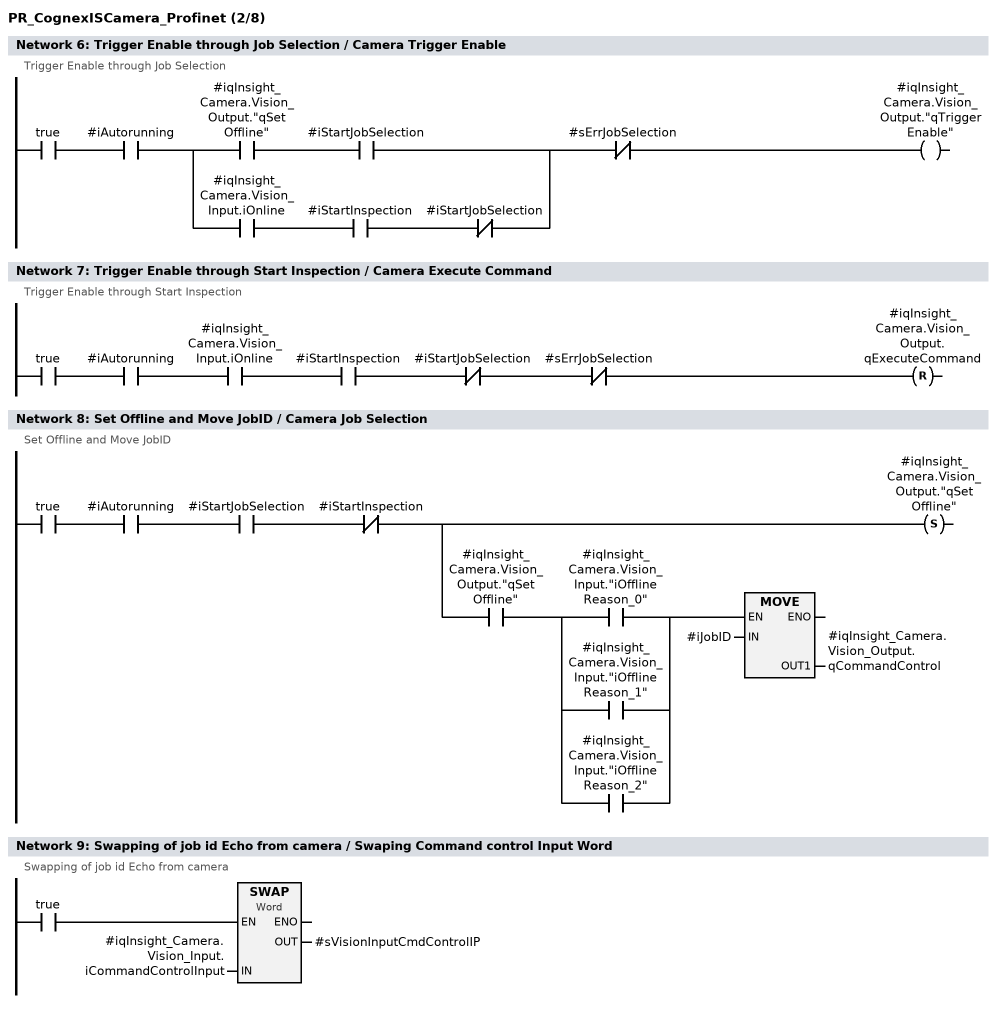
   RUNG wire#powerrail
      Contact( true )
      Contact( #iAutorunning )
      wire#w1
      Contact( #iqInsight_Camera.Vision_Output."qSet Offline" )
      Contact( #iStartJobSelection )
      wire#w2
      I_Contact( #sErrJobSelection )
      Coil( #iqInsight_Camera.Vision_Output."qTrigger Enable" )
   END_RUNG
   RUNG wire#w1
      Contact( #iqInsight_Camera.Vision_Input.iOnline )
      Contact( #iStartInspection )
      I_Contact( #iStartJobSelection )
   END_RUNG wire#w2
   // the same network as SCL:
   #iqInsight_Camera.Vision_Output."qTrigger Enable" := true AND #iAutorunning AND ((#iqInsight_Camera.Vision_Output."qSet Offline" AND #iStartJobSelection) OR (#iqInsight_Camera.Vision_Input.iOnline AND #iStartInspection AND NOT #iStartJobSelection)) AND NOT #sErrJobSelection;
END_REGION

REGION Network 7: Trigger Enable through Start Inspection / Camera Execute Command
   // Trigger Enable through Start Inspection
   RUNG wire#powerrail
      Contact( true )
      Contact( #iAutorunning )
      Contact( #iqInsight_Camera.Vision_Input.iOnline )
      Contact( #iStartInspection )
      I_Contact( #iStartJobSelection )
      I_Contact( #sErrJobSelection )
      R_Coil( #iqInsight_Camera.Vision_Output.qExecuteCommand )
   END_RUNG
   // the same network as SCL:
   IF true AND #iAutorunning AND #iqInsight_Camera.Vision_Input.iOnline AND #iStartInspection AND NOT #iStartJobSelection AND NOT #sErrJobSelection THEN
       #iqInsight_Camera.Vision_Output.qExecuteCommand := FALSE;
   END_IF;
END_REGION

REGION Network 8: Set Offline and Move JobID / Camera Job Selection
   // Set Offline and Move JobID
   RUNG wire#powerrail
      Contact( true )
      Contact( #iAutorunning )
      Contact( #iStartJobSelection )
      I_Contact( #iStartInspection )
      wire#w1
      S_Coil( #iqInsight_Camera.Vision_Output."qSet Offline" )
   END_RUNG
   RUNG wire#w1
      Contact( #iqInsight_Camera.Vision_Output."qSet Offline" )
      wire#w2
      Contact( #iqInsight_Camera.Vision_Input."iOffline Reason_0" )
      wire#w3
      Move(in := #iJobID, out1 => #iqInsight_Camera.Vision_Output.qCommandControl)
   END_RUNG
   RUNG wire#w2
      Contact( #iqInsight_Camera.Vision_Input."iOffline Reason_1" )
   END_RUNG wire#w3
   RUNG wire#w2
      Contact( #iqInsight_Camera.Vision_Input."iOffline Reason_2" )
   END_RUNG wire#w3
   // the same network as SCL:
   #_w1 := true AND #iAutorunning AND #iStartJobSelection AND NOT #iStartInspection;
   IF #_w1 THEN #iqInsight_Camera.Vision_Output."qSet Offline" := TRUE; END_IF;
   IF #_w1 AND #iqInsight_Camera.Vision_Output."qSet Offline" AND (#iqInsight_Camera.Vision_Input."iOffline Reason_0" OR #iqInsight_Camera.Vision_Input."iOffline Reason_1" OR #iqInsight_Camera.Vision_Input."iOffline Reason_2") THEN
       #iqInsight_Camera.Vision_Output.qCommandControl := #iJobID;
   END_IF;
END_REGION

REGION Network 9: Swapping of job id Echo from camera / Swaping Command control Input Word
   // Swapping of job id Echo from camera
   IF true THEN
       #sVisionInputCmdControlIP := SWAP(#iqInsight_Camera.Vision_Input.iCommandControlInput);
   END_IF;
END_REGION

REGION Network 10: Initiate Job Load / Camera Execute Command
   // Initiate Job Load
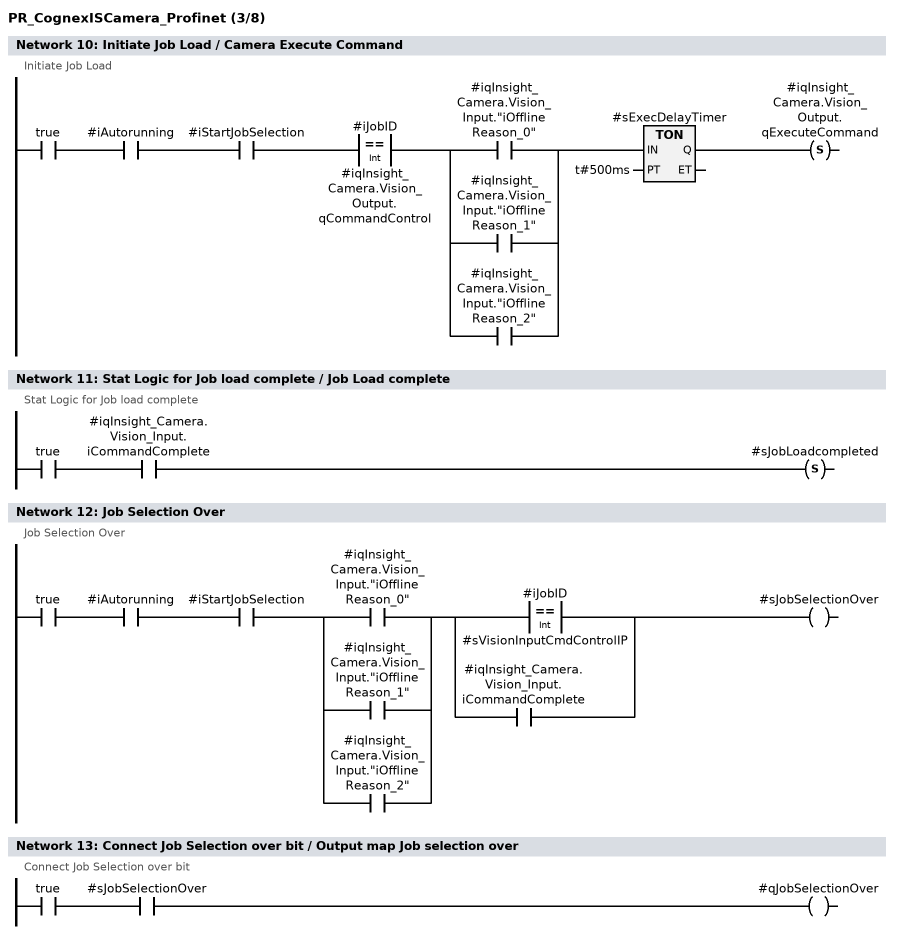
   #sExecDelayTimer(IN := true AND #iAutorunning AND #iStartJobSelection AND (#iJobID = #iqInsight_Camera.Vision_Output.qCommandControl) AND (#iqInsight_Camera.Vision_Input."iOffline Reason_0" OR #iqInsight_Camera.Vision_Input."iOffline Reason_1" OR #iqInsight_Camera.Vision_Input."iOffline Reason_2"),   // TON
                    PT := t#500ms);
   IF #sExecDelayTimer.Q THEN #iqInsight_Camera.Vision_Output.qExecuteCommand := TRUE; END_IF;
END_REGION

REGION Network 11: Stat Logic for Job load complete / Job Load complete
   // Stat Logic for Job load complete
   RUNG wire#powerrail
      Contact( true )
      Contact( #iqInsight_Camera.Vision_Input.iCommandComplete )
      S_Coil( #sJobLoadcompleted )
   END_RUNG
   // the same network as SCL:
   IF true AND #iqInsight_Camera.Vision_Input.iCommandComplete THEN #sJobLoadcompleted := TRUE; END_IF;
END_REGION

REGION Network 12: Job Selection Over
   // Job Selection Over
   RUNG wire#powerrail
      Contact( true )
      Contact( #iAutorunning )
      Contact( #iStartJobSelection )
      wire#w1
      Contact( #iqInsight_Camera.Vision_Input."iOffline Reason_0" )
      wire#w2
      { S7_Templates := "SrcType := Int" } EQ_Contact(in1 := #iJobID, in2 := #sVisionInputCmdControlIP)
      wire#w3
      Coil( #sJobSelectionOver )
   END_RUNG
   RUNG wire#w1
      Contact( #iqInsight_Camera.Vision_Input."iOffline Reason_1" )
   END_RUNG wire#w2
   RUNG wire#w1
      Contact( #iqInsight_Camera.Vision_Input."iOffline Reason_2" )
   END_RUNG wire#w2
   RUNG wire#w2
      Contact( #iqInsight_Camera.Vision_Input.iCommandComplete )
   END_RUNG wire#w3
   // the same network as SCL:
   #sJobSelectionOver := true AND #iAutorunning AND #iStartJobSelection AND (#iqInsight_Camera.Vision_Input."iOffline Reason_0" OR #iqInsight_Camera.Vision_Input."iOffline Reason_1" OR #iqInsight_Camera.Vision_Input."iOffline Reason_2") AND ((#iJobID = #sVisionInputCmdControlIP) OR #iqInsight_Camera.Vision_Input.iCommandComplete);
END_REGION

REGION Network 13: Connect Job Selection over bit / Output map Job selection over
   // Connect Job Selection over bit
   RUNG wire#powerrail
      Contact( true )
      Contact( #sJobSelectionOver )
      Coil( #qJobSelectionOver )
   END_RUNG
   // the same network as SCL:
   #qJobSelectionOver := true AND #sJobSelectionOver;
END_REGION

REGION Network 14: Reset Offline / Camera Job Selection reset
   // Reset Offline / "#iqInsight_Camera.Vision_Output.qSet Offline" and "#iqInsight_Camera.Vision_Output.qExecuteCommand"  Reset coil removed while block comparision
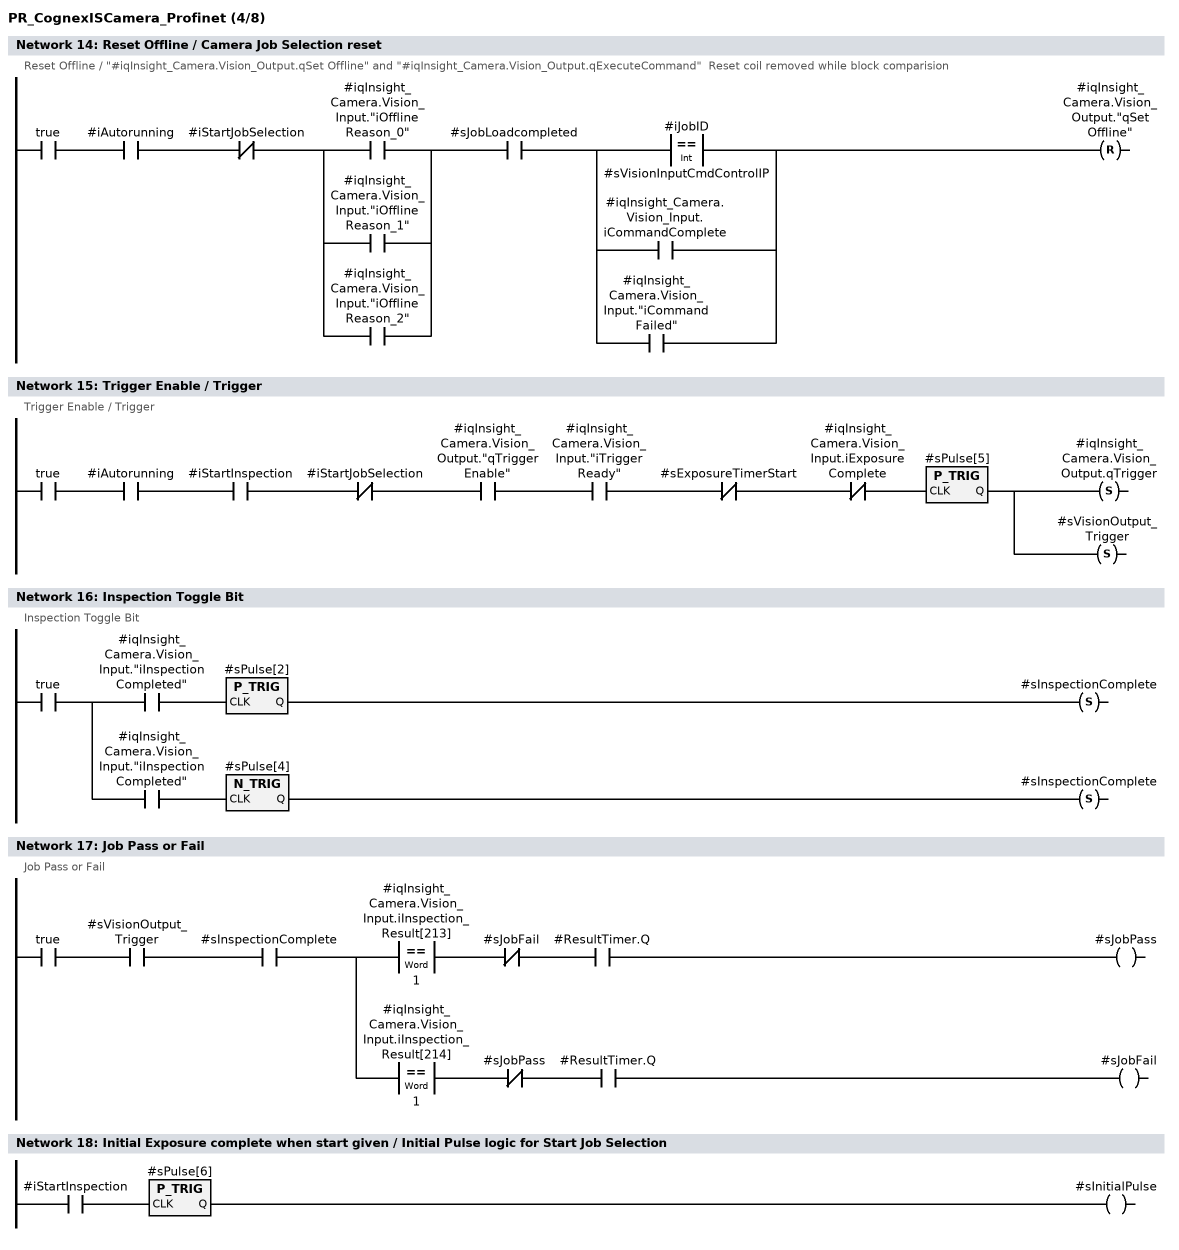
   RUNG wire#powerrail
      Contact( true )
      Contact( #iAutorunning )
      I_Contact( #iStartJobSelection )
      wire#w1
      Contact( #iqInsight_Camera.Vision_Input."iOffline Reason_0" )
      wire#w2
      Contact( #sJobLoadcompleted )
      wire#w3
      { S7_Templates := "SrcType := Int" } EQ_Contact(in1 := #iJobID, in2 := #sVisionInputCmdControlIP)
      wire#w4
      R_Coil( #iqInsight_Camera.Vision_Output."qSet Offline" )
   END_RUNG
   RUNG wire#w1
      Contact( #iqInsight_Camera.Vision_Input."iOffline Reason_1" )
   END_RUNG wire#w2
   RUNG wire#w1
      Contact( #iqInsight_Camera.Vision_Input."iOffline Reason_2" )
   END_RUNG wire#w2
   RUNG wire#w3
      Contact( #iqInsight_Camera.Vision_Input.iCommandComplete )
   END_RUNG wire#w4
   RUNG wire#w3
      Contact( #iqInsight_Camera.Vision_Input."iCommand Failed" )
   END_RUNG wire#w4
   // the same network as SCL:
   IF true AND #iAutorunning AND NOT #iStartJobSelection AND (#iqInsight_Camera.Vision_Input."iOffline Reason_0" OR #iqInsight_Camera.Vision_Input."iOffline Reason_1" OR #iqInsight_Camera.Vision_Input."iOffline Reason_2") AND #sJobLoadcompleted AND ((#iJobID = #sVisionInputCmdControlIP) OR #iqInsight_Camera.Vision_Input.iCommandComplete OR #iqInsight_Camera.Vision_Input."iCommand Failed") THEN
       #iqInsight_Camera.Vision_Output."qSet Offline" := FALSE;
   END_IF;
END_REGION

REGION Network 15: Trigger Enable / Trigger
   // Trigger Enable / Trigger
   RUNG wire#powerrail
      Contact( true )
      Contact( #iAutorunning )
      Contact( #iStartInspection )
      I_Contact( #iStartJobSelection )
      Contact( #iqInsight_Camera.Vision_Output."qTrigger Enable" )
      Contact( #iqInsight_Camera.Vision_Input."iTrigger Ready" )
      I_Contact( #sExposureTimerStart )
      I_Contact( #iqInsight_Camera.Vision_Input.iExposureComplete )
      P_Trig( #sPulse[5] )
      wire#w1
      S_Coil( #iqInsight_Camera.Vision_Output.qTrigger )
   END_RUNG
   RUNG wire#w1
      S_Coil( #sVisionOutput_Trigger )
   END_RUNG
   // the same network as SCL:
   #_w1 := true AND #iAutorunning AND #iStartInspection AND NOT #iStartJobSelection AND #iqInsight_Camera.Vision_Output."qTrigger Enable" AND #iqInsight_Camera.Vision_Input."iTrigger Ready" AND NOT #sExposureTimerStart AND NOT #iqInsight_Camera.Vision_Input.iExposureComplete;
   #_w2 := #_w1 AND NOT #sPulse[5];   // rising edge
   #sPulse[5] := #_w1;
   IF #_w2 THEN
       #iqInsight_Camera.Vision_Output.qTrigger := TRUE;
       #sVisionOutput_Trigger := TRUE;
   END_IF;
END_REGION

REGION Network 16: Inspection Toggle Bit
   // Inspection Toggle Bit
   RUNG wire#powerrail
      Contact( true )
      wire#w1
      Contact( #iqInsight_Camera.Vision_Input."iInspection Completed" )
      P_Trig( #sPulse[2] )
      S_Coil( #sInspectionComplete )
   END_RUNG
   RUNG wire#w1
      Contact( #iqInsight_Camera.Vision_Input."iInspection Completed" )
      N_Trig( #sPulse[4] )
      S_Coil( #sInspectionComplete )
   END_RUNG
   // the same network as SCL:
   #_w1 := true AND #iqInsight_Camera.Vision_Input."iInspection Completed";
   #_w2 := #_w1 AND NOT #sPulse[2];   // rising edge
   #sPulse[2] := #_w1;
   IF #_w2 THEN #sInspectionComplete := TRUE; END_IF;
   #_w3 := true AND #iqInsight_Camera.Vision_Input."iInspection Completed";
   #_w4 := NOT #_w3 AND #sPulse[4];   // falling edge
   #sPulse[4] := #_w3;
   IF #_w4 THEN #sInspectionComplete := TRUE; END_IF;
END_REGION

REGION Network 17: Job Pass or Fail
   // Job Pass or Fail
   RUNG wire#powerrail
      Contact( true )
      Contact( #sVisionOutput_Trigger )
      Contact( #sInspectionComplete )
      wire#w1
      { S7_Templates := "SrcType := Word" } EQ_Contact(in1 := #iqInsight_Camera.Vision_Input.iInspection_Result[213], in2 := 1)
      I_Contact( #sJobFail )
      Contact( #ResultTimer.Q )
      Coil( #sJobPass )
   END_RUNG
   RUNG wire#w1
      { S7_Templates := "SrcType := Word" } EQ_Contact(in1 := #iqInsight_Camera.Vision_Input.iInspection_Result[214], in2 := 1)
      I_Contact( #sJobPass )
      Contact( #ResultTimer.Q )
      Coil( #sJobFail )
   END_RUNG
   // the same network as SCL:
   #_w1 := true AND #sVisionOutput_Trigger AND #sInspectionComplete;
   #sJobPass := #_w1 AND (#iqInsight_Camera.Vision_Input.iInspection_Result[213] = 1) AND NOT #sJobFail AND #ResultTimer.Q;
   #sJobFail := #_w1 AND (#iqInsight_Camera.Vision_Input.iInspection_Result[214] = 1) AND NOT #sJobPass AND #ResultTimer.Q;
END_REGION

REGION Network 18: Initial Exposure complete when start given / Initial Pulse logic for Start Job Selection
   RUNG wire#powerrail
      Contact( #iStartInspection )
      P_Trig( #sPulse[6] )
      Coil( #sInitialPulse )
   END_RUNG
   // the same network as SCL:
   #_w1 := #iStartInspection AND NOT #sPulse[6];   // rising edge
   #sPulse[6] := #iStartInspection;
   #sInitialPulse := #_w1;
END_REGION

REGION Network 19: Exposure Timer 1
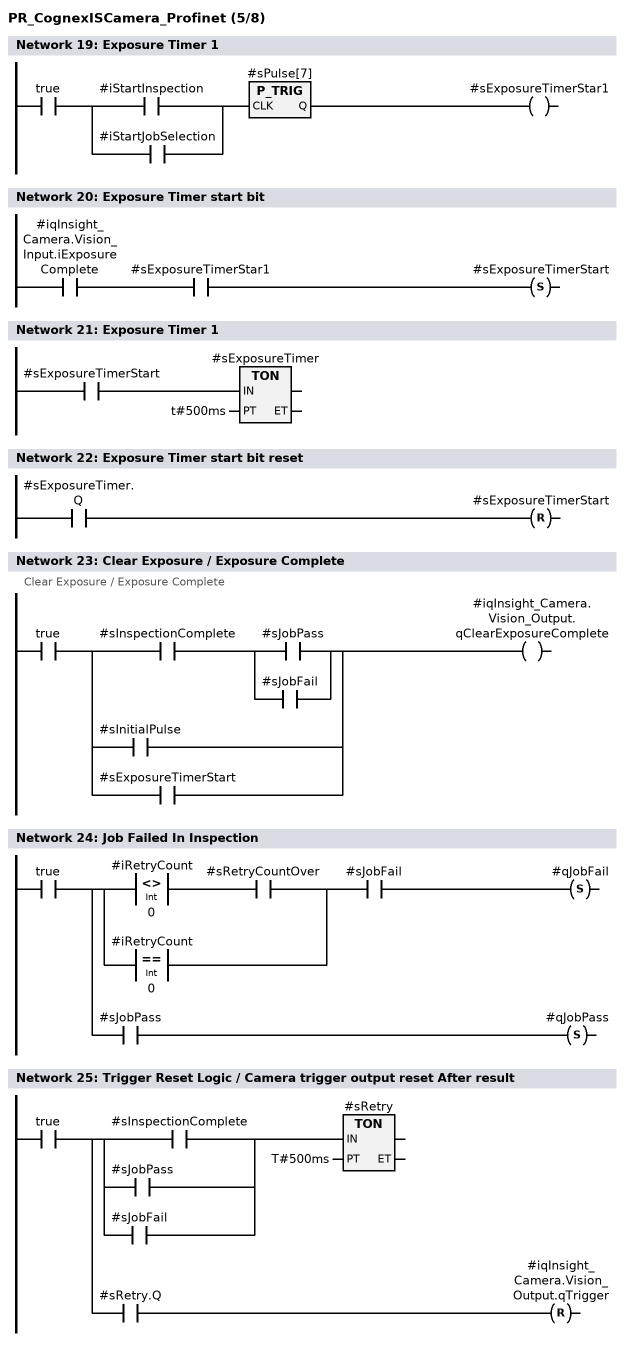
   RUNG wire#powerrail
      Contact( true )
      wire#w1
      Contact( #iStartInspection )
      wire#w2
      P_Trig( #sPulse[7] )
      Coil( #sExposureTimerStar1 )
   END_RUNG
   RUNG wire#w1
      Contact( #iStartJobSelection )
   END_RUNG wire#w2
   // the same network as SCL:
   #_w1 := true AND (#iStartInspection OR #iStartJobSelection);
   #_w2 := #_w1 AND NOT #sPulse[7];   // rising edge
   #sPulse[7] := #_w1;
   #sExposureTimerStar1 := #_w2;
END_REGION

REGION Network 20: Exposure Timer start bit
   RUNG wire#powerrail
      Contact( #iqInsight_Camera.Vision_Input.iExposureComplete )
      Contact( #sExposureTimerStar1 )
      S_Coil( #sExposureTimerStart )
   END_RUNG
   // the same network as SCL:
   IF #iqInsight_Camera.Vision_Input.iExposureComplete AND #sExposureTimerStar1 THEN
       #sExposureTimerStart := TRUE;
   END_IF;
END_REGION

REGION Network 21: Exposure Timer 1
   #sExposureTimer(IN := #sExposureTimerStart, PT := t#500ms);   // TON
END_REGION

REGION Network 22: Exposure Timer start bit reset
   RUNG wire#powerrail
      Contact( #sExposureTimer.Q )
      R_Coil( #sExposureTimerStart )
   END_RUNG
   // the same network as SCL:
   IF #sExposureTimer.Q THEN #sExposureTimerStart := FALSE; END_IF;
END_REGION

REGION Network 23: Clear Exposure / Exposure Complete
   // Clear Exposure / Exposure Complete
   RUNG wire#powerrail
      Contact( true )
      wire#w1
      Contact( #sInspectionComplete )
      wire#w2
      Contact( #sJobPass )
      wire#w3
      Coil( #iqInsight_Camera.Vision_Output.qClearExposureComplete )
   END_RUNG
   RUNG wire#w2
      Contact( #sJobFail )
   END_RUNG wire#w3
   RUNG wire#w1
      Contact( #sInitialPulse )
   END_RUNG wire#w3
   RUNG wire#w1
      Contact( #sExposureTimerStart )
   END_RUNG wire#w3
   // the same network as SCL:
   #iqInsight_Camera.Vision_Output.qClearExposureComplete := true AND ((#sInspectionComplete AND (#sJobPass OR #sJobFail)) OR #sInitialPulse OR #sExposureTimerStart);
END_REGION

REGION Network 24: Job Failed In Inspection
   RUNG wire#powerrail
      Contact( true )
      wire#w1
      { S7_Templates := "SrcType := Int" } NE_Contact(in1 := #iRetryCount, in2 := 0)
      Contact( #sRetryCountOver )
      wire#w2
      Contact( #sJobFail )
      S_Coil( #qJobFail )
   END_RUNG
   RUNG wire#w1
      { S7_Templates := "SrcType := Int" } EQ_Contact(in1 := #iRetryCount, in2 := 0)
   END_RUNG wire#w2
   RUNG wire#w1
      Contact( #sJobPass )
      S_Coil( #qJobPass )
   END_RUNG
   // the same network as SCL:
   IF true AND (((#iRetryCount <> 0) AND #sRetryCountOver) OR (#iRetryCount = 0)) AND #sJobFail THEN
       #qJobFail := TRUE;
   END_IF;
   IF true AND #sJobPass THEN #qJobPass := TRUE; END_IF;
END_REGION

REGION Network 25: Trigger Reset Logic / Camera trigger output reset After result
   #sRetry(IN := true AND (#sInspectionComplete OR #sJobPass OR #sJobFail), PT := T#500ms);   // TON
   IF true AND #sRetry.Q THEN #iqInsight_Camera.Vision_Output.qTrigger := FALSE; END_IF;
END_REGION

REGION Network 26: Retry Count Logic / CameraTrigger Enable on for retry count
   // Retry Count Logic
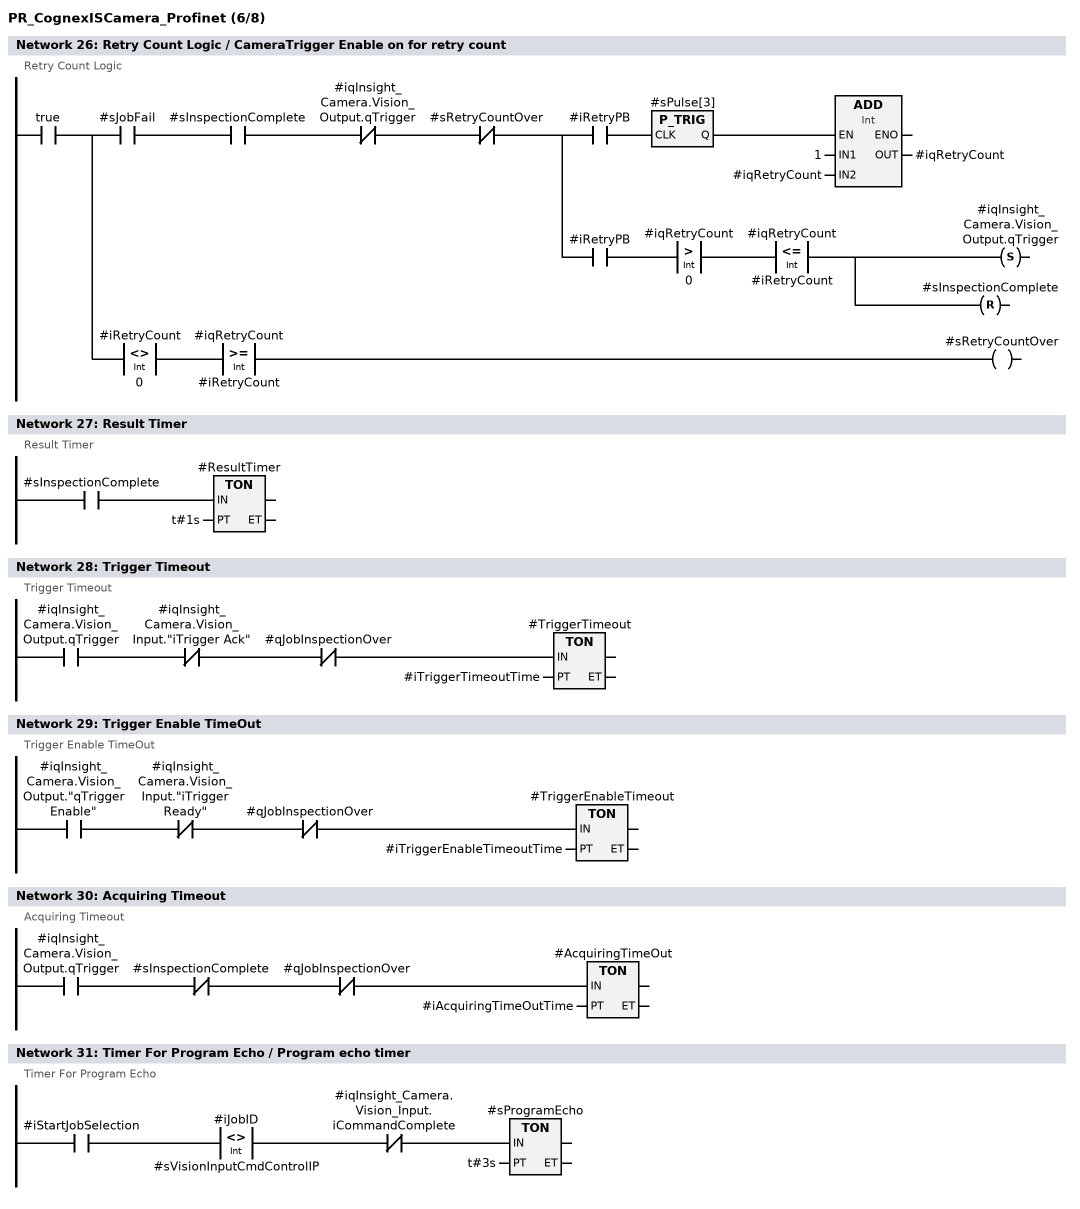
   RUNG wire#powerrail
      Contact( true )
      wire#w1
      Contact( #sJobFail )
      Contact( #sInspectionComplete )
      I_Contact( #iqInsight_Camera.Vision_Output.qTrigger )
      I_Contact( #sRetryCountOver )
      wire#w2
      Contact( #iRetryPB )
      P_Trig( #sPulse[3] )
      { S7_Templates := "SrcType := Int" } Add(in1 := 1, in2 := #iqRetryCount, out => #iqRetryCount)
   END_RUNG
   RUNG wire#w2
      Contact( #iRetryPB )
      { S7_Templates := "SrcType := Int" } GT_Contact(in1 := #iqRetryCount, in2 := 0)
      { S7_Templates := "SrcType := Int" } LE_Contact(in1 := #iqRetryCount, in2 := #iRetryCount)
      wire#w3
      S_Coil( #iqInsight_Camera.Vision_Output.qTrigger )
   END_RUNG
   RUNG wire#w3
      R_Coil( #sInspectionComplete )
   END_RUNG
   RUNG wire#w1
      { S7_Templates := "SrcType := Int" } NE_Contact(in1 := #iRetryCount, in2 := 0)
      { S7_Templates := "SrcType := Int" } GE_Contact(in1 := #iqRetryCount, in2 := #iRetryCount)
      Coil( #sRetryCountOver )
   END_RUNG
   // the same network as SCL:
   #_w1 := true AND #sJobFail AND #sInspectionComplete AND NOT #iqInsight_Camera.Vision_Output.qTrigger AND NOT #sRetryCountOver;
   #_w2 := #_w1 AND #iRetryPB;
   #_w3 := #_w2 AND NOT #sPulse[3];   // rising edge
   #sPulse[3] := #_w2;
   IF #_w3 THEN #iqRetryCount := 1 + #iqRetryCount; END_IF;
   IF #_w1 AND #iRetryPB AND (#iqRetryCount > 0) AND (#iqRetryCount <= #iRetryCount) THEN
       #iqInsight_Camera.Vision_Output.qTrigger := TRUE;
       #sInspectionComplete := FALSE;
   END_IF;
   #sRetryCountOver := true AND (#iRetryCount <> 0) AND (#iqRetryCount >= #iRetryCount);
END_REGION

REGION Network 27: Result Timer
   // Result Timer
   #ResultTimer(IN := #sInspectionComplete, PT := t#1s);   // TON
END_REGION

REGION Network 28: Trigger Timeout
   // Trigger Timeout
   #TriggerTimeout(IN := #iqInsight_Camera.Vision_Output.qTrigger AND NOT #iqInsight_Camera.Vision_Input."iTrigger Ack" AND NOT #qJobInspectionOver,   // TON
                   PT := #iTriggerTimeoutTime);
END_REGION

REGION Network 29: Trigger Enable TimeOut
   // Trigger Enable TimeOut
   #TriggerEnableTimeout(IN := #iqInsight_Camera.Vision_Output."qTrigger Enable" AND NOT #iqInsight_Camera.Vision_Input."iTrigger Ready" AND NOT #qJobInspectionOver,   // TON
                         PT := #iTriggerEnableTimeoutTime);
END_REGION

REGION Network 30: Acquiring Timeout
   // Acquiring Timeout
   #AcquiringTimeOut(IN := #iqInsight_Camera.Vision_Output.qTrigger AND NOT #sInspectionComplete AND NOT #qJobInspectionOver,   // TON
                     PT := #iAcquiringTimeOutTime);
END_REGION

REGION Network 31: Timer For Program Echo / Program echo timer
   // Timer For Program Echo
   #sProgramEcho(IN := #iStartJobSelection AND (#iJobID <> #sVisionInputCmdControlIP) AND NOT #iqInsight_Camera.Vision_Input.iCommandComplete,   // TON
                 PT := t#3s);
END_REGION

REGION Network 32: OutPuts
   // OutPuts
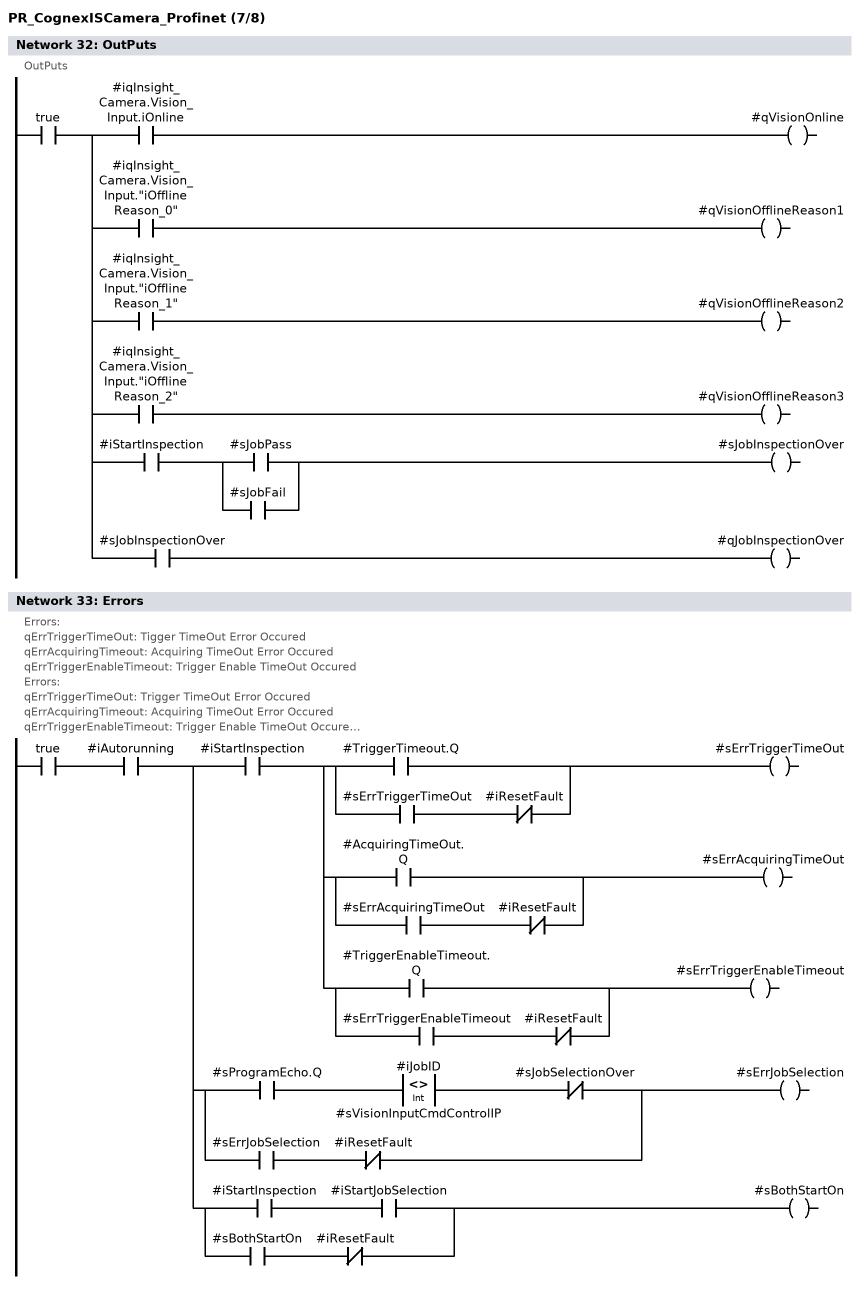
   RUNG wire#powerrail
      Contact( true )
      wire#w1
      Contact( #iqInsight_Camera.Vision_Input.iOnline )
      Coil( #qVisionOnline )
   END_RUNG
   RUNG wire#w1
      Contact( #iqInsight_Camera.Vision_Input."iOffline Reason_0" )
      Coil( #qVisionOfflineReason1 )
   END_RUNG
   RUNG wire#w1
      Contact( #iqInsight_Camera.Vision_Input."iOffline Reason_1" )
      Coil( #qVisionOfflineReason2 )
   END_RUNG
   RUNG wire#w1
      Contact( #iqInsight_Camera.Vision_Input."iOffline Reason_2" )
      Coil( #qVisionOfflineReason3 )
   END_RUNG
   RUNG wire#w1
      Contact( #iStartInspection )
      wire#w2
      Contact( #sJobPass )
      wire#w3
      Coil( #sJobInspectionOver )
   END_RUNG
   RUNG wire#w2
      Contact( #sJobFail )
   END_RUNG wire#w3
   RUNG wire#w1
      Contact( #sJobInspectionOver )
      Coil( #qJobInspectionOver )
   END_RUNG
   // the same network as SCL:
   #qVisionOnline := true AND #iqInsight_Camera.Vision_Input.iOnline;
   #qVisionOfflineReason1 := true AND #iqInsight_Camera.Vision_Input."iOffline Reason_0";
   #qVisionOfflineReason2 := true AND #iqInsight_Camera.Vision_Input."iOffline Reason_1";
   #qVisionOfflineReason3 := true AND #iqInsight_Camera.Vision_Input."iOffline Reason_2";
   #sJobInspectionOver := true AND #iStartInspection AND (#sJobPass OR #sJobFail);
   #qJobInspectionOver := true AND #sJobInspectionOver;
END_REGION

REGION Network 33: Errors
   // Errors: 
   // qErrTriggerTimeOut: Tigger TimeOut Error Occured
   // qErrAcquiringTimeout: Acquiring TimeOut Error Occured
   // qErrTriggerEnableTimeout: Trigger Enable TimeOut Occured
   // Errors: 
   // qErrTriggerTimeOut: Trigger TimeOut Error Occured
   // qErrAcquiringTimeout: Acquiring TimeOut Error Occured
   // qErrTriggerEnableTimeout: Trigger Enable TimeOut Occured
   // qErrJobSelection: Job selection Error
   // qBothStartOn: Both Start are ON
   RUNG wire#powerrail
      Contact( true )
      Contact( #iAutorunning )
      wire#w1
      Contact( #iStartInspection )
      wire#w2
      Contact( #TriggerTimeout.Q )
      wire#w3
      Coil( #sErrTriggerTimeOut )
   END_RUNG
   RUNG wire#w2
      Contact( #sErrTriggerTimeOut )
      I_Contact( #iResetFault )
   END_RUNG wire#w3
   RUNG wire#w2
      Contact( #AcquiringTimeOut.Q )
      wire#w4
      Coil( #sErrAcquiringTimeOut )
   END_RUNG
   RUNG wire#w2
      Contact( #sErrAcquiringTimeOut )
      I_Contact( #iResetFault )
   END_RUNG wire#w4
   RUNG wire#w2
      Contact( #TriggerEnableTimeout.Q )
      wire#w5
      Coil( #sErrTriggerEnableTimeout )
   END_RUNG
   RUNG wire#w2
      Contact( #sErrTriggerEnableTimeout )
      I_Contact( #iResetFault )
   END_RUNG wire#w5
   RUNG wire#w1
      Contact( #sProgramEcho.Q )
      { S7_Templates := "SrcType := Int" } NE_Contact(in1 := #iJobID, in2 := #sVisionInputCmdControlIP)
      I_Contact( #sJobSelectionOver )
      wire#w6
      Coil( #sErrJobSelection )
   END_RUNG
   RUNG wire#w1
      Contact( #sErrJobSelection )
      I_Contact( #iResetFault )
   END_RUNG wire#w6
   RUNG wire#w1
      Contact( #iStartInspection )
      Contact( #iStartJobSelection )
      wire#w7
      Coil( #sBothStartOn )
   END_RUNG
   RUNG wire#w1
      Contact( #sBothStartOn )
      I_Contact( #iResetFault )
   END_RUNG wire#w7
   // the same network as SCL:
   #_w1 := true AND #iAutorunning;
   #_w2 := #_w1 AND #iStartInspection;
   #sErrTriggerTimeOut := #_w2 AND (#TriggerTimeout.Q OR (#sErrTriggerTimeOut AND NOT #iResetFault));
   #sErrAcquiringTimeOut := #_w2 AND (#AcquiringTimeOut.Q OR (#sErrAcquiringTimeOut AND NOT #iResetFault));
   #sErrTriggerEnableTimeout := #_w2 AND (#TriggerEnableTimeout.Q OR (#sErrTriggerEnableTimeout AND NOT #iResetFault));
   #sErrJobSelection := #_w1 AND ((#sProgramEcho.Q AND (#iJobID <> #sVisionInputCmdControlIP) AND NOT #sJobSelectionOver) OR (#sErrJobSelection AND NOT #iResetFault));
   #sBothStartOn := #_w1 AND ((#iStartInspection AND #iStartJobSelection) OR (#sBothStartOn AND NOT #iResetFault));
END_REGION

REGION Network 34: Stat bit Error Mapping / Output mapping using Stat Bit
   // Stat bit Error Mapping / Output mapping using Stat Bit
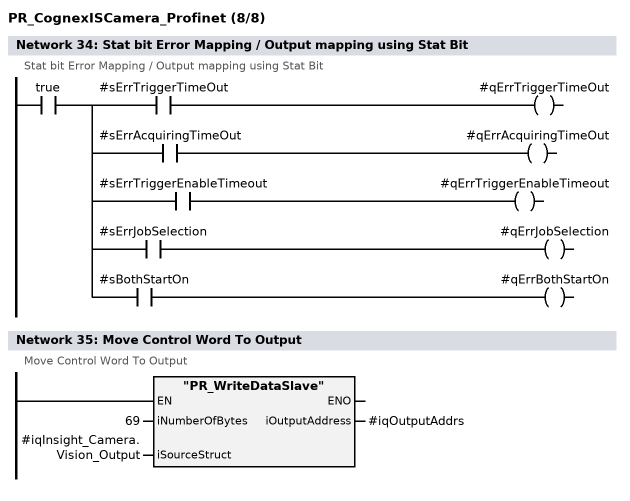
   RUNG wire#powerrail
      Contact( true )
      wire#w1
      Contact( #sErrTriggerTimeOut )
      Coil( #qErrTriggerTimeOut )
   END_RUNG
   RUNG wire#w1
      Contact( #sErrAcquiringTimeOut )
      Coil( #qErrAcquiringTimeOut )
   END_RUNG
   RUNG wire#w1
      Contact( #sErrTriggerEnableTimeout )
      Coil( #qErrTriggerEnableTimeout )
   END_RUNG
   RUNG wire#w1
      Contact( #sErrJobSelection )
      Coil( #qErrJobSelection )
   END_RUNG
   RUNG wire#w1
      Contact( #sBothStartOn )
      Coil( #qErrBothStartOn )
   END_RUNG
   // the same network as SCL:
   #qErrTriggerTimeOut := true AND #sErrTriggerTimeOut;
   #qErrAcquiringTimeOut := true AND #sErrAcquiringTimeOut;
   #qErrTriggerEnableTimeout := true AND #sErrTriggerEnableTimeout;
   #qErrJobSelection := true AND #sErrJobSelection;
   #qErrBothStartOn := true AND #sBothStartOn;
END_REGION

REGION Network 35: Move Control Word To Output
   // Move Control Word To Output
   RUNG wire#powerrail
      "PR_WriteDataSlave"(iNumberOfBytes := 69, iSourceStruct := #iqInsight_Camera.Vision_Output, iOutputAddress => #iqOutputAddrs)
   END_RUNG
   // the same network as SCL:
   "PR_WriteDataSlave"(iNumberOfBytes := 69,
                       iSourceStruct := #iqInsight_Camera.Vision_Output,
                       iOutputAddress => #iqOutputAddrs);
END_REGION
END_FUNCTION_BLOCK

FUNCTION_BLOCK "PR_CognexIS28xx_Profi"   // FB496, LAD
TITLE = PR_CognexIS28xx_Profi
{ S7_Optimized_Access := 'TRUE' }
AUTHOR : MS
FAMILY : WiproPari
NAME : S21006022015
VERSION : 0.3
   VAR_INPUT
      iInsightCamera_Input : "UDT_IS28xx_To_Plc";   // Connect Camera Input
      iResetFault : Bool;   // Reset Fault Input
      iModuleReset : Bool;   // Connect Module reset Signal to this pin
      iAutorunning : Bool;   // Autorunning Input
      iStartJobSelection : Bool;   // start job selection
      iStartInspection : Bool;   // start inspection
      iJobID : Int;   // job id
      iUserData : Array[1..60] of Byte;   // Enter user data which is send to cognex camera/controller
      iTriggerEnableTimeoutTime : Time;   // Trigger Enable TimeOut Time Delay
      iTriggerTimeoutTime : Time;   // Trigger TimeOut Time Delay
      iAcquiringTimeOutTime : Time;   // Acquiring TimeOut Time Delay
      iPrgmNoTimeOut : Time;   // Timeout for program echo received from camera
      iFeedbackTimeOut : Time;   // Feedback time out time
   END_VAR
   VAR_OUTPUT
      qInsightCamera_Output : "UDT_Plc_To_IS28xx";   // Connect Camera Output
      qJobPass : Bool;   // Job Pass In Inspection
      qJobFail : Bool;   // Job Failed In Inspection
      qJobSelectionOver : Bool;   // job selection over
      qJobInspectionOver : Bool;   // Inspection Over Output
      qVisionOnline : Bool;   // Insight Vision Is In Online
      qVisionOfflineReason1 : Bool;   // Insight Vision Offline Due To: The vision system's job is being modified
      qVisionOfflineReason2 : Bool;   // Insight Vision Offline Due To: A discrete signal is holding the vision system Offline
      qVisionOfflineReason3 : Bool;   // Insight Vision Offline Due To: A communications protocol is holding the vision system Offline
      qErrBothStartOn : Bool;   // both start on
      qErrJobSelection : Bool;   // error job selection
      qErrTriggerEnableTimeout : Bool;   // Trigger Enable TimeOut Error
      qErrTriggerTimeOut : Bool;   // Trigger TimeOut Error
      qErrAcquiringTimeOut : Bool;   // Acquiring TimeOut Error
      qErrJobIDEchoMismatch : Bool;   // Job Id Echo mismatch Error
      qErrSetUserDataAckNtRcvd : Bool;   // Set user data ack not received within time
      qMsgJobIDMismatch : Bool;   // Selected Job ID & Running JOB ID not matched message
      qInspectionResult : Array[1..60] of Byte;   // Inspection Result Data
   END_VAR
   VAR_IN_OUT
      iqRunningJobID : Int;   // It Shows running Job ID
   END_VAR
   VAR
      sResetFaults : Bool;
      sInspectionComplete : Bool;
      sJobPass : Bool;
      sJobFail : Bool;
      sJobLoadcompleted : Bool;
      sJobSelectionOver : Bool;
      sJobInspectionOver : Bool;
      sVisionOutput_Trigger : Bool;
      sInitialPulse : Bool;
      sExposureTimerStar1 : Bool;
      sExposureTimerStart : Bool;
      sPulse : Array[0..7] of Bool;
      sVisionInputCmdControlIP : Int;
      sTriggerEnableTimeoutTime : Time;
      sTriggerTimeoutTime : Time;
      sAcquiringTimeOutTime : Time;
      TriggerTimeout : TON_TIME;
      TriggerEnableTimeout : TON_TIME;
      AcquiringTimeOut : TON_TIME;
      ResultTimer : TON_TIME;
      sExposureTimer : TON_TIME;
      sTriggerResetTimer : TON_TIME;
      sPrgmNoTimeOut : Time;
      sPrgmNumTimer : TON_TIME;
      sSetUserDataAckTimer : TON_TIME;
      sFeedbackTimeOut : Time;
   END_VAR
   VAR_TEMP   // added for the SCL form of the ladder/FBD networks
      _w1 : Bool;
      _w2 : Bool;
      _w3 : Bool;
      _w4 : Bool;
      _w5 : Bool;
   END_VAR
BEGIN

